  def limit(value, range):
      return scale(value, range, range)
  end


  rq_init_comm_if_connected(9, "1")
  rq_init_comm_if_connected(2, "2")
  rq_init_comm_if_connected(3, "3")
  rq_init_comm_if_connected(4, "4")
  rq_print_connected_grippers()
  rq_gripper_communication_thread = run rq_gripper_communication()
  set_closed_norm(97.6470588235294, 1)
  set_open_norm(1.1764705882352942, 1)
  set_closed_mm(0.0, 1)
  set_open_mm(53.0, 1)
  set_closed_norm(100.0, 2)
  set_open_norm(0.0, 2)
  set_closed_mm(0.0, 2)
  set_open_mm(50.0, 2)
  set_closed_norm(100.0, 3)
  set_open_norm(0.0, 3)
  set_closed_mm(0.0, 3)
  set_open_mm(50.0, 3)
  set_closed_norm(100.0, 4)
  set_open_norm(0.0, 4)
  set_closed_mm(0.0, 4)
  set_open_mm(50.0, 4)
  rq_current_limit_enabled = False
  while(not rq_gripper_communication_thread_started):
      sync()
  end
  # end: URCap Installation Node
  # begin: URCap Installation Node
  #   Source: OPC UA, 2.0.2, Rocketfarm AS
  #   Type: OPC UA
  global opcua_daemon = rpc_factory("xmlrpc", "http://127.0.0.1:40409/RPC2")
  def opcua_client_connect(address):
  return opcua_daemon.client_connect(address)
  end
  def opcua_client_get_id(client_name):
  return opcua_daemon.client_get_id(client_name)
  end
  def opcua_client_try_connect(client_id):
  opcua_result = False
  if (opcua_daemon.client_connect(client_id)):
  sleep(0.01)
  opcua_result = opcua_daemon.client_is_connected(client_id)
  opcua_retry = 10
  while ( (not opcua_result) and (opcua_retry > 0) ):
  sleep(0.1)
  opcua_result = opcua_daemon.client_is_connected(client_id)
  opcua_retry = opcua_retry - 1
  end
  end
  return opcua_result
  end
  def opcua_client_disconnect(client_id):
  return opcua_daemon.client_disconnect(client_id)
  end
  def opcua_client_is_connected(client_id):
  return opcua_daemon.client_is_connected(client_id)
  end
  def opcua_client_read_byid(client_id, namespace_id, variable_id):
  return opcua_daemon.client_read_variable_by_id(client_id, namespace_id, variable_id)
  end
  def opcua_client_read_byname(client_id, namespace_id, variable_name):
  return opcua_daemon.client_read_variable_by_name(client_id, namespace_id, variable_name)
  end
  def opcua_client_write_byid(client_id, namespace_id, variable_id, variable_value):
  return opcua_daemon.client_write_variable_by_id(client_id, namespace_id, variable_id, variable_value)
  end
  def opcua_client_write_byname(client_id, namespace_id, variable_name, variable_value):
  return opcua_daemon.client_write_variable_by_name(client_id, namespace_id, variable_name, variable_value)
  end
  def opcua_client_last_error(client_id):
  return opcua_daemon.client_get_last_error(client_id)
  end
  def opcua_server_read_byname(variable_name):
  return opcua_daemon.server_read_variable_by_name(variable_name)
  end
  def opcua_server_write_byname(variable_name, variable_value):
  return opcua_daemon.server_write_variable_by_name(variable_name, variable_value)
  end
  def opcua_server_last_error():
  return opcua_daemon.server_get_last_error()
  end
  def opcua_error_to_string(errorCode):
  return opcua_daemon.error_code_to_string(errorCode)
  end
  # end: URCap Installation Node
  step_count_7be696b6_0fa4_4b27_b09b_633ea860953e = 0.0
  thread Step_Counter_Thread_93e352b0_e34b_423c_bc3a_28ecb8afdc0a():
    while (True):
      step_count_7be696b6_0fa4_4b27_b09b_633ea860953e = step_count_7be696b6_0fa4_4b27_b09b_633ea860953e + 1.0
      sync()
    end
  end
  run Step_Counter_Thread_93e352b0_e34b_423c_bc3a_28ecb8afdc0a()
  global AMR_Position=struct(position_identifier=0, x1=0, x2=0, y1=0, y2=0, theta1=0, theta2=0)
  global CAM_Pose=p[0,0,0,0,0,0]
  global CAM_Relation=""
  global CMD_Abort=  False
  global CMD_Clear=  False
  global CMD_Reset=  False
  global CMD_Start=  False
  global CMD_Suspend=  False
  global CMD_Unhold=  False
  global CMD_Unsuspend=  False
  global CNT_Rack_Output=0
  global FNC_Freedrive=  False
  global PRC_TubCounter=0
  global PRC_TubNumber=0
  global STP=0
  global easyPickCount=0
  global easyPickCount_5=0
  global easyPickNoObj=0
  global easyPickNoObj_5=0
  global easyPickParts=0
  global easyPickParts_5=0
  global TMR_Barcode=0
  global Container_mid_1_p=p[-.379239199143, -.127191311915, .299999999998, .000000000046, -.000000000021, -1.247199999994]
  global Container_mid_1_q=[-2.477408934449926, -1.2969853503591224, -1.875639182904262, -1.539621866126728, 1.5731943360401213, -2.8009955944022717]
  global Container_capt_p=p[-.525590029047, .407247642794, .411588185841, -.000000000107, .000000000065, -2.896148821900]
  global Container_capt_q=[-3.5968351615224767, -2.0050156108707204, -0.8176271154495112, -1.8895759482008394, 1.5730967555598792, -2.2743681102957645]
  global Waypoint_6_p=p[.008800512419, -.547926542621, .402696567415, -.589884378425, -.007228654778, -.061268144704]
  global Waypoint_6_q=[-1.2044575850116175, -1.3416667741588135, -1.8272563219070435, -0.9884541195682068, 1.3621035814285278, -2.7712565104113978]
  global Waypoint_18_p=p[-.178371829612, -.433927395311, .368082383916, -.086593488055, .704679941724, -.007869906074]
  global Waypoint_18_q=[-1.265390698109762, -1.3355963987163086, -1.7944865226745605, -1.7402602634825648, 0.8780410885810852, -2.7713127771960657]
  global Waypoint_12_p=p[.008800512419, -.547926542621, .402696567415, -.589884378425, -.007228654778, -.061268144704]
  global Waypoint_12_q=[-1.2044575850116175, -1.3416667741588135, -1.8272563219070435, -0.9884541195682068, 1.3621035814285278, -2.7712565104113978]
  global Waypoint_19_p=p[-.178371829612, -.433927395311, .368082383916, -.086593488055, .704679941724, -.007869906074]
  global Waypoint_19_q=[-1.265390698109762, -1.3355963987163086, -1.7944865226745605, -1.7402602634825648, 0.8780410885810852, -2.7713127771960657]
  global Vial_above_p=p[.017105793010, -.652093028359, .184920586844, .000000000272, .000000000270, 1.564063451276]
  global Vial_above_q=[-1.3375440709712851, -1.9618096977868804, -1.4665759083780685, -1.2837941559171444, 1.5732503672317195, -4.47276330421513]
  global Vial_pick_point_p=p[.017105792852, -.648922724010, .093307568731, .000000000271, .000000000270, 1.564063451276]
  global Vial_pick_point_q=[-1.3366329456391917, -2.0375277831965413, -1.6071432798879028, -1.0675084332049813, 1.57309887265915, -4.471135348858068]
  global Waypoint_20_p=p[.019227646885, -.648669633640, .184920586950, .000000000000, .000000000000, .024063451426]
  global Waypoint_20_q=[-1.3331129109407733, -1.9540750545686123, -1.4775914902901128, -1.280581784992414, 1.5733500744865856, -2.928303704452631]
  global Waypoint_33_p=p[-.032361834699, -.348336136197, .391475576335, -.000008499254, .000014589902, -.004651426820]
  global Waypoint_33_q=[-1.2709335019096129, -1.1914598663441005, -1.708995335060501, -1.8117888533498316, 1.5729683532263925, -2.8379347397710237]
  global Vial_3FG_place_p=p[-.031858676359, -.349402499566, .145301120695, .000000000000, .000000000000, .000000000000]
  global Vial_3FG_place_q=[-1.2723975525801707, -1.252376585823825, -2.3128114007049496, -1.1470592278900167, 1.5730548099411423, -2.8414815174610535]
  global Waypoint_34_p=p[-.032361834699, -.348336136197, .391475576335, -.000008499254, .000014589902, -.004651426820]
  global Waypoint_34_q=[-1.2709335019096129, -1.1914598663441005, -1.708995335060501, -1.8117888533498316, 1.5729683532263925, -2.8379347397710237]
  global cap_dump_p=p[-.139168676487, -.420163541420, .146096395183, .000000000000, .000000000000, .000000000000]
  global cap_dump_q=[-1.584588644510994, -1.5093464179777323, -2.1118449369620347, -1.091059703602438, 1.5728943834877336, -3.154014906686923]
  global Waypoint_35_p=p[-.032361834699, -.348336136197, .391475576335, -.000008499254, .000014589902, -.004651426820]
  global Waypoint_35_q=[-1.2709335019096129, -1.1914598663441005, -1.708995335060501, -1.8117888533498316, 1.5729683532263925, -2.8379347397710237]
  global Waypoint_36_p=p[-.032361834699, -.348336136197, .391475576335, -.000008499254, .000014589902, -.004651426820]
  global Waypoint_36_q=[-1.2709335019096129, -1.1914598663441005, -1.708995335060501, -1.8117888533498316, 1.5729683532263925, -2.8379347397710237]
  global Waypoint_37_p=p[-.032361834699, -.348336136197, .391475576335, -.000008499254, .000014589902, -.004651426820]
  global Waypoint_37_q=[-1.2709335019096129, -1.1914598663441005, -1.708995335060501, -1.8117888533498316, 1.5729683532263925, -2.8379347397710237]
  global Vial_liq_above_p=p[-.025303660977, -.338758622354, .426628485936, -1.315858642253, .800043520260, -.928295855026]
  global Vial_liq_above_q=[-0.3789628187762659, -1.5149522957256814, -2.263045310974121, 0.7870649534412841, -0.750984017048971, -3.2237566153155726]
  global Vial_liq_pick_1_p=p[-.002660428945, -.335984893034, .159389832934, -1.150456778400, .673175527684, -1.010612657503]
  global Vial_liq_pick_1_q=[-0.3660772482501429, -1.4503649038127442, -2.4056053161621094, -1.994692941705221, 0.8039668202400208, -0.2508929411517542]
  global Vial_liq_pick_2_p=p[-.041402486291, -.356791603314, .125395323246, -1.143483969075, .651070210027, -.878721885453]
  global Vial_liq_pick_2_q=[-0.4426233705502476, -1.437252121513727, -2.551930962114307, -1.776528229806984, 0.6562026234073748, -0.43018811960029524]
  global Liquid_midway_p=p[.057575295009, -.583081747994, .306414980749, -1.351675548728, .120935756539, -.096908606303]
  global Liquid_midway_q=[-0.895174805318014, -1.7035466633238734, -2.380953073501587, 0.631549521083496, 0.7706599235534668, -2.9455552736865442]
  global shake_1_p=p[.057574880217, -.583085370269, .306422893466, -1.360996190983, -.155555042453, -.438136255921]
  global shake_1_q=[-0.8951800505267542, -1.7035466633238734, -2.380937099456787, 0.6315542894550782, 0.7706599235534669, -2.5394540616517496]
  global shake_2_p=p[.057581636113, -.583090570002, .306439684073, -1.308767904323, .368530312677, .214926493520]
  global shake_2_q=[-0.8951714674579065, -1.7035395107665003, -2.380906343460083, 0.6315504747578125, 0.7706480026245118, -3.3161255787892268]
  global drop_above_1_p=p[.268235025993, -.467784390499, .226219872376, -1.027832627524, -.430841408251, 1.004603115937]
  global drop_above_1_q=[-0.935645882283346, -1.6663371525206507, -2.4252893924713135, 0.41966931402172847, 1.8470635414123535, -3.4600217978106897]
  global drop_above_2_p=p[.219042229014, -.470775657081, .133754190740, -.313004595901, -.344395319364, 1.500564994056]
  global drop_above_2_q=[-1.0601594887284795, -1.70046459045642, -2.0799996233759863, -0.7243227230676759, 1.9429634314685202, -4.115129153870795]
  global liq_tran_1_p=p[.213067510942, -.469567035397, .100231043184, .251862243732, .217902579404, 1.592812335393]
  global liq_tran_1_q=[-0.7789645168037476, -1.822364827406652, -1.8643518410805573, -1.252158963840138, 1.3768134449520435, -3.9328333233290254]
  global Waypoint_21_p=p[.187119460405, -.493959476151, .133754190608, -.313004596540, -.344395317757, 1.500564993991]
  global Waypoint_21_q=[-1.1418328121400876, -1.7310553375189475, -2.033634768766424, -0.772026910513711, 1.958578934631971, -4.201588449364511]
  global liq_tran_2_p=p[.195957706507, -.493022614126, .100231042689, .160718757180, .109807038912, 1.525321508623]
  global liq_tran_2_q=[-0.881740380645474, -1.8244526267589851, -1.865100964490387, -1.1608866323693583, 1.4631433601076713, -3.973915130363038]
  global Vial_drop_above_p=p[.000324902251, -.648569523142, .221894115667, -.873462921366, 1.165852672573, -1.482720593185]
  global Vial_drop_above_q=[-1.0576906334721352, -2.393016994184633, -0.9236232851859159, -2.5729213042279273, 0.7903331288549689, -0.33286325848155585]
  global Vial_liq_drop_p=p[.001020867953, -.647659915585, .092915870838, -.834762611599, 1.081942994823, -1.540647900176]
  global Vial_liq_drop_q=[-1.0631954168193474, -2.4447642951220825, -1.128811017825127, -2.1983115491972294, 0.8130148661460634, -0.38984988696911316]
  global Waypoint_9_p=p[.206300564882, -.401796282405, .209941275233, .000000000049, .000000000063, 1.560839127857]
  global Waypoint_9_q=[-0.7963359454512808, -1.4686025034365713, -1.9726632321075135, -1.2709582822971974, 1.5730203818053559, -3.9272300959189193]
  global Waypoint_10_p=p[.200865824304, -.400817692024, .105072686738, .000000000049, .000000000061, 1.560839127855]
  global Waypoint_10_q=[-0.8042914374275529, -1.5824702465090397, -2.1630314773482997, -0.9667217216455377, 1.5726337265768082, -3.9342465798801403]
  global Waypoint_11_p=p[.200865824280, -.400817691999, .325177251663, .000000000049, .000000000061, 1.560839127855]
  global Waypoint_11_q=[-0.8031609769098491, -1.4190566846320642, -1.7173307870816634, -1.5758364190022327, 1.5730457436482617, -3.935202548332848]
  global Waypoint_7_p=p[-.615828862681, .233809157513, .299999999960, .005115849907, .008741794022, -2.111813105778]
  global Waypoint_7_q=[-3.2957401409809868, -1.9361965884744503, -1.2056078493731617, -1.569266158150004, 1.5650998100608482, -2.7562028470627613]
  global Waypoint_8_p=p[-.615828862366, .233809157463, .013910424379, .005115849905, .008741794020, -2.111813105780]
  global Waypoint_8_q=[-3.2964782505943173, -2.1586184138220776, -1.6500090431308791, -0.9024541777239836, 1.5648120752692236, -2.7547026290098384]
  global Waypoint_13_p=p[-.479450777041, .284140798427, .125270103493, -.276792173670, 2.098433187455, -2.121256516887]
  global Waypoint_13_q=[-2.8915050665484827, -1.9549266300597132, -2.2318272590637207, -1.6654960117735804, 0.020810842514038086, -0.4019392172442835]
  global Waypoint_70_p=p[-.472820924464, .292439826304, .207418370234, -.259787347864, -2.053484648504, 2.070709755662]
  global Waypoint_70_q=[-2.969927421603815, -2.07168115810532, -1.6835546062719366, -2.4953958198513964, 0.4489790927922641, -0.005578998612037367]
  global Waypoint_1_p=p[-.312961047461, -.152991312519, .223609826854, -.745314530454, -1.713873240489, 1.673341715282]
  global Waypoint_1_q=[-2.3560472170459192, -2.183784624139303, -1.4583134651184082, -2.6435262165465296, 1.6522362232208252, 0.043451953679323196]
  global Waypoint_16_p=p[-.113749865836, -.390110151572, .317307487562, -.519383711706, -.839884211339, 1.756868173041]
  global Waypoint_16_q=[-1.8909733931170862, -1.720626016656393, -1.5115610361099243, -2.1240560017027796, 2.1809096336364746, 0.7227501273155212]
  global Waypoint_15_p=p[.029144035010, -.436802470887, .327885032028, -.521560953301, -.623641814548, 1.862659450154]
  global Waypoint_15_q=[-1.564817253743307, -1.556895188321807, -1.6826975345611572, -1.6944714985289515, 2.2362685203552246, 1.117417335510254]
  global Waypoint_14_p=p[.068712235638, -.569419545175, .285215357659, -.679242949116, -.712065334485, 1.394044574094]
  global Waypoint_14_q=[-1.5731792953485346, -1.8029235103747094, -1.6781008808776736, -1.2218450646111982, 2.4719572998240125, 1.6394218026856375]
  global Waypoint_17_p=p[-.047220457210, -.557624911767, .136370962514, -.679242949107, -.712065334475, 1.394044574096]
  global Waypoint_17_q=[-1.7740079055958748, -2.0023561428872334, -1.7577251142892676, -1.18903287716154, 2.4487287370345143, 1.322902469273079]
  global Waypoint_25_p=p[.065436479647, -.569388431626, .287820755049, -.679242949185, -.712065334557, 1.394044574070]
  global Waypoint_25_q=[-1.5789263550890595, -1.8020194754825436, -1.6702557537748035, -1.237882536889547, 2.471995808083492, 1.6301087487321393]
  global Waypoint_73_p=p[.200650292861, -.570238752026, .330084459991, 1.360500825815, .021700154388, 2.681649888469]
  global Waypoint_73_q=[-0.7671117850166942, -2.170180210127774, -0.8654875324671831, -2.4760661058854714, 1.019668964673781, 1.1886838746103445]
  global Waypoint_51_p=p[.143029822311, -.569853361759, .275754213782, 1.297896664289, .026410127072, 2.712872144875]
  global Waypoint_51_q=[-0.8339941389801577, -2.0499669090260237, -1.181859109742545, -2.1992567984298894, 0.9933974691724003, 1.1053015960835664]
  global Waypoint_55_p=p[.073857253409, -.577012553496, .221504790513, 1.297896665457, .026410123899, 2.712872144362]
  global Waypoint_55_q=[-0.9235026509638331, -2.0031911550113533, -1.4013130080059835, -1.9791459123699324, 0.9364696407276547, 1.0224867664664226]
  global Waypoint_56_p=p[.135677267144, -.579447716527, .242231366835, 1.555421348248, .015405426287, 2.555899922373]
  global Waypoint_56_q=[-0.8277598345563266, -2.1783820448240228, -1.1390951780517948, -2.3437042464770936, 0.9222576608739947, 1.2572681804986878]
  global Waypoint_57_p=p[.143391004007, -.581808738942, .226065325532, 1.639743959545, .007914821713, 2.502360786858]
  global Waypoint_57_q=[-0.8163397121067408, -2.2409861865625498, -1.1056400409378426, -2.4000192569642436, 0.9131014133193622, 1.3141118037187605]
  global Waypoint_59_p=p[.272401132286, -.578182925380, .239561357365, 2.126997331910, .113921148153, 2.155615020515]
  global Waypoint_59_q=[-0.6600120703326624, -2.700596948663229, -0.4450863301753998, -3.1158048115172328, 0.9327830672264099, 1.686402678489685]
  global Waypoint_58_p=p[.223648508176, -.578477552733, .276546452136, 2.174288010107, -.044108754041, 2.058653287678]
  global Waypoint_58_q=[-0.7290484882560344, -2.6749849159411134, -0.44426632073579775, -3.220833992584847, 0.9665895014735898, 1.686536774549042]
  global Waypoint_60_p=p[-.013316432876, -.544772031582, .383371643081, 2.208233379808, .037543335712, 2.097559881761]
  global Waypoint_60_q=[-0.9328326161883087, -2.0999933666355775, -1.1958015693111372, -3.060905141293654, 0.690378518537611, 1.7121940951337198]
  global Waypoint_61_p=p[-.412188693372, -.356446875193, .383371643081, 1.751740964455, -.739956256289, 1.600691174920]
  global Waypoint_61_q=[-1.766185342973321, -2.0999933666355775, -1.1958015693111372, -3.060905141293654, 0.690378518537611, 1.7121940951337198]
  global Waypoint_62_p=p[-.542658707241, -.114281911009, .251261544113, 1.813043609523, -.679411528034, 1.655271622964]
  global Waypoint_62_q=[-2.158300033470912, -1.9418836862428677, -1.8142999147147894, -2.778920736683023, 0.21900622104017292, 1.8983390235012934]
  global Waypoint_63_p=p[-.532496162227, -.127810170801, .159342327524, 1.813043609478, -.679411528027, 1.655271622994]
  global Waypoint_63_q=[-2.1232624524640213, -2.086114053133292, -1.8911847933380095, -2.5248779786918614, 0.2536249317365024, 1.864405460969639]
  global Waypoint_52_p=p[-.576034890047, -.066269986912, .306739617770, .862065193359, -.255405331227, 2.195240951653]
  global Waypoint_52_q=[-2.4808268779922003, -1.5303848711262056, -1.876845562237385, -1.1257011427858359, 0.8740163290385958, -0.15002503295170655]
  global Waypoint_69_p=p[-.581965326699, -.059291422286, .312082125679, .862065195757, -.255405329473, 2.195240950921]
  global Waypoint_69_q=[-2.500621389999687, -1.5361955180345959, -1.8614018767844556, -1.1190332887072278, 0.8777181708365909, -0.17540933674578696]
  global Waypoint_71_p=p[-.581965326670, -.059291422265, .290575803625, .862065195756, -.255405329472, 2.195240950921]
  global Waypoint_71_q=[-2.5007210652259566, -1.5510704265538795, -1.9040561970342402, -1.0615823481403304, 0.8776641555740685, -0.17528706367848557]
  global Waypoint_72_p=p[-.581965326627, -.059291422244, .350142125738, 1.757497900770, -.677813691618, 1.696469016977]
  global Waypoint_72_q=[-2.3014470577960933, -1.774776476208789, -1.7081605706825291, -2.8433626113276596, 0.07508598567825443, 1.682946898281932]
  global Waypoint_68_p=p[-.333292906431, -.480744165508, .350142125738, 2.217519979286, .140864133573, 2.209123277630]
  global Waypoint_68_q=[-1.438387057796029, -1.774776476208789, -1.7081605706825291, -2.8433626113276596, 0.07508598567825443, 1.682946898281932]
  global TMR_Barcode_is_counting=False
  thread Timer_Thread():
    while (True):
      if (TMR_Barcode_is_counting):
        TMR_Barcode = TMR_Barcode + get_steptime()
      end
      sync()
    end
  end
  run Timer_Thread()
  def Sub_Vision_V18():
    $ 697 "Sub_Vision_V18" "noBreak"
    $ 698 "PreSettings"
    $ 699 "CAM_LM_Detected≔ False "
    global CAM_LM_Detected=  False
    $ 700 "CAM_Captures≔0"
    global CAM_Captures=0
    $ 701 "CAM_Pose≔p[0,0,0,0,0,0]"
    global CAM_Pose=p[0,0,0,0,0,0]
    $ 702 "CAM_LM_Refinmnt≔ False "
    global CAM_LM_Refinmnt=  False
    $ 703 "CAM_LM_Refined≔ False "
    global CAM_LM_Refined=  False
    $ 704 "CAM_LM_Deviatn≔p[0,0,0,0,0,0]"
    global CAM_LM_Deviatn=p[0,0,0,0,0,0]
    $ 705 "CAM_LM_ID≔0"
    global CAM_LM_ID=0
    $ 706 "CAM_Done≔ False "
    global CAM_Done=  False
    $ 707 "CAM_CNT_Obj≔0"
    global CAM_CNT_Obj=0
    $ 708 "CAM_Result = []"
    CAM_Result = []
    $ 709 "OBJ_Detected≔ False "
    global OBJ_Detected=  False
    $ 710 "FRM_Reference≔p[0,0,0,0,0,0]"
    global FRM_Reference=p[0,0,0,0,0,0]
    $ 711 "'=========='"
    # '=========='
    $ 712 "Switch Action"
    switch_1 = Action
    $ 713 "Case 13"
    if (13 == switch_1):
    elif (15 == switch_1):
      $ 831 "Case 15"
    elif (131 == switch_1):
      $ 877 "Case 131"
      $ 878 "Read (SensoPart)"
      $ 879 "Action_Info≔'search for landmark'"
      global Action_Info="search for landmark"
      $ 880 "CAM_LM≔CAM_LMs[4]"
      global CAM_LM=CAM_LMs[4]
      $ 881 "CAM_Relation≔CAM_LM.capture_relation"
      global CAM_Relation=CAM_LM.capture_relation
      $ 882 "go to capture pose"
      $ 885 "If ITM_ID≟1 and JIG≟7"
      if (ITM_ID == 1  and  JIG == 7):
        $ 886 "PSE_T≔uLM_Cap_SSRack"
        global PSE_T=uLM_Cap_SSRack
      else:
        $ 887 "ElseIf ITM_ID≟5 and JIG≟7"
        if (ITM_ID == 5  and  JIG == 7):
          $ 888 "PSE_T≔FRM_Cap_SSRack"
          global PSE_T=FRM_Cap_SSRack
        else:
          $ 889 "ElseIf ITM_ID≟13 and JIG≟7"
          if (ITM_ID == 13  and  JIG == 7):
            $ 890 "PSE_T≔FRM_pick_rack_const"
            global PSE_T=p[-0.5568395192387274,0.34423986364170267,0.44698620470146266,-1.0069110132199915E-6,3.378712467497258E-5,-8.002029546773325E-6]
          else:
            $ 891 "ElseIf ITM_ID≟1 and JIG≟15"
            if (ITM_ID == 1 and JIG == 15):
              $ 892 "MoveJ"
              $ 893 "Container_mid_1" "breakAfter"
              movej(get_inverse_kin(Container_mid_1_p, qnear=Container_mid_1_q), a=1.3962634015954636, v=1.0471975511965976, r=0.05)
              $ 894 "Container_capt" "breakAfter"
              movej(get_inverse_kin(Container_capt_p, qnear=Container_capt_q), a=1.3962634015954636, v=1.0471975511965976)
              $ 895 "PSE_T≔FRM_Container_S_const"
              global PSE_T=p[-0.510412665574981,0.40064363362973565,0.41159789496794374,-1.1370875604168537E-5,-3.643547521609506E-6,-2.896122366208473]
            end
          end
        end
      end
      $ 896 "do_transition(PSE_T, keep_rxry=False)"
      do_transition(PSE_T, keep_rxry=False)
      $ 897 "Set"
      set_tcp(p[0.0,0.0,0.161,3.1415,0.0,0.0])
      $ 898 "MoveJ"
      $ 899 "PSE_T" "breakAfter"
      movej(PSE_T, a=1.3962634015954636, v=1.7453292519943295)
      $ 900 "CAM_Pose≔get_actual_tcp_pose()"
      global CAM_Pose= get_actual_tcp_pose ()
      $ 901 "Loop  not CAM_Done and  not ERROR.FLAG and  not CMD_Stop"
      while (  not  CAM_Done  and    not  ERROR.FLAG  and    not  CMD_Stop):
        $ 902 "adjust capture pose"
        $ 903 "If CAM_LM_Detected and CAM_LM_Refinmnt"
        if (CAM_LM_Detected  and  CAM_LM_Refinmnt):
          $ 904 "PSE_T≔p[0,0,0.300,0,0,0]"
          global PSE_T=p[0,0,0.300,0,0,0]
          $ 905 "CAM_Pose≔PSE_T"
          global CAM_Pose=PSE_T
          $ 906 "If  not is_reachable(FRM_Reference,[PSE_T])"
          if (  not  is_reachable(FRM_Reference,[PSE_T])):
            $ 907 "Error"
            $ 908 "set_error(ERROR_POSE_NOT_REACHABLE)"
            set_error(ERROR_POSE_NOT_REACHABLE)
          end
          $ 909 "If  not ERROR.FLAG"
          if (  not  ERROR.FLAG):
            $ 910 "MoveJ"
            $ 911 "PSE_T" "breakAfter"
            set_tcp(p[0.0,0.0,0.161,0.0,0.0,0.0])
            movej(pose_trans(FRM_Reference, PSE_T), a=0.8726646259971648, v=1.3962634015954636)
            $ 912 "CAM_LM_Refined≔ True "
            global CAM_LM_Refined=  True
          end
        else:
          $ 913 "ElseIf  not CAM_LM_Detected and CAM_Captures>0"
          if (  not  CAM_LM_Detected  and  CAM_Captures>0):
            $ 914 "MoveL"
            $ 915 "If FRM_Reference≟p[0,0,0,0,0,0]"
            if (FRM_Reference == p[0,0,0,0,0,0]):
              $ 916 "PSE_T≔get_random_pose(pose_ref=CAM_Pose, mode='cubic', range_max=[0.150,0.150,0.015])"
              global PSE_T=get_random_pose(pose_ref=CAM_Pose, mode="cubic", range_max=[0.150,0.150,0.015])
            else:
              $ 921 "Else" "noBreak"
              $ 922 "PSE_T≔get_random_pose(pose_ref=CAM_Pose, mode='rotation', range_max=[10,10,0])"
              global PSE_T=get_random_pose(pose_ref=CAM_Pose, mode="rotation", range_max=[10,10,0])
              $ 923 "CAM_LM_Refined≔ True "
              global CAM_LM_Refined=  True
            end
            $ 924 "If get_inverse_kin_has_solution(pose_trans(FRM_Reference, PSE_T))"
            if (get_inverse_kin_has_solution( pose_trans (FRM_Reference, PSE_T))):
              $ 925 "Comment"
              # Comment
              $ 926 "PSE_T" "breakAfter"
              set_tcp(p[0.0,0.0,0.161,3.1415,0.0,0.0])
              movel(pose_trans(FRM_Reference, PSE_T), a=0.03, v=0.05)
            else:
              $ 927 "Else" "noBreak"
              $ 928 "'If random pose is out of reach, set the initial cam pose'"
              # 'If random pose is out of reach, set the initial cam pose'
              $ 929 "PSE_T≔CAM_Pose"
              global PSE_T=CAM_Pose
            end
          end
        end
        $ 930 "Wait: 2.0"
        sleep(2.0)
        $ 931 "trigger"
        $ 932 "If ITM_ID≟1 and JIG≟7"
        if (ITM_ID == 1  and  JIG == 7):
          # begin: URCap Program Node
          #   Source: SensoPart VISOR Robotic, 2.0.0, SensoPart Industriesensorik GmbH
          #   Type: VISOR Trigger
          $ 933 "# 1 VISOR Trigger"
          visor_changeJob(1, "Landmark_INVITE_2", 6000)
          visor_trigger(1, 6000, "arm")
          # end: URCap Program Node
        else:
          $ 934 "ElseIf ITM_ID≟5 and JIG≟7"
          if (ITM_ID == 5  and  JIG == 7):
            # begin: URCap Program Node
            #   Source: SensoPart VISOR Robotic, 2.0.0, SensoPart Industriesensorik GmbH
            #   Type: VISOR Trigger
            $ 935 "# 1 VISOR Trigger"
            visor_changeJob(1, "Landmark_INVITE_2", 6000)
            visor_trigger(1, 6000, "arm")
            # end: URCap Program Node
          else:
            $ 936 "ElseIf ITM_ID≟13 and JIG≟7"
            if (ITM_ID == 13  and  JIG == 7):
              # begin: URCap Program Node
              #   Source: SensoPart VISOR Robotic, 2.0.0, SensoPart Industriesensorik GmbH
              #   Type: VISOR Trigger
              $ 937 "# 1 VISOR Trigger"
              visor_changeJob(1, "Landmark_INVITE_2", 6000)
              visor_trigger(1, 6000, "arm")
              # end: URCap Program Node
            else:
              $ 938 "ElseIf ITM_ID≟1 and JIG≟15"
              if (ITM_ID == 1 and JIG == 15):
                # begin: URCap Program Node
                #   Source: SensoPart VISOR Robotic, 2.0.0, SensoPart Industriesensorik GmbH
                #   Type: VISOR Trigger
                $ 939 "# 1 VISOR Trigger"
                visor_changeJob(1, "Container_S", 6000)
                visor_trigger(1, 6000, "arm")
                # end: URCap Program Node
              end
            end
          end
        end
        $ 943 "TM_3D_Found≔visor_partsFound(1)"
        global TM_3D_Found= visor_partsFound (1)
        $ 944 "If TM_3D_Found>0"
        if (TM_3D_Found>0):
          $ 945 "CAM_LM_Detected≔ True "
          global CAM_LM_Detected=  True
          $ 946 "CAM_Captures≔0"
          global CAM_Captures=0
        else:
          $ 947 "Else" "noBreak"
          $ 948 "CAM_LM_Detected≔ False "
          global CAM_LM_Detected=  False
          $ 949 "CAM_Captures≔CAM_Captures+1"
          global CAM_Captures=CAM_Captures+1
        end
        $ 954 "result"
        $ 955 "If CAM_LM_Detected"
        if (CAM_LM_Detected):
          $ 956 "If (CAM_LM_Refinmnt and CAM_LM_Refined) or  not CAM_LM_Refinmnt"
          if ((CAM_LM_Refinmnt  and  CAM_LM_Refined)  or    not  CAM_LM_Refinmnt):
            $ 1014 "If ITM_ID≟1 and JIG≟7"
            if (ITM_ID == 1  and  JIG == 7):
              $ 1015 "CAM_LM_SSRack≔visor_getPose3d(1, 0)"
              global CAM_LM_SSRack= visor_getPose3d (1, 0)
            else:
              $ 1016 "ElseIf ITM_ID≟5 and JIG≟7"
              if (ITM_ID == 5  and  JIG == 7):
                $ 1017 "CAM_LM_SSRack≔visor_getPose3d(1, 0)"
                global CAM_LM_SSRack= visor_getPose3d (1, 0)
              else:
                $ 1018 "ElseIf ITM_ID≟13 and JIG≟7"
                if (ITM_ID == 13  and  JIG == 7):
                  $ 1019 "CAM_LM_Bott≔visor_getPose3d(1, 0)"
                  global CAM_LM_Bott= visor_getPose3d (1, 0)
                else:
                  $ 1020 "ElseIf ITM_ID≟1 and JIG≟15"
                  if (ITM_ID == 1 and JIG == 15):
                    $ 1021 "CAM_LM_Cont_S≔visor_getPose3d(1, 0)"
                    global CAM_LM_Cont_S= visor_getPose3d (1, 0)
                  end
                end
              end
            end
            $ 1022 "CAM_Done≔ True "
            global CAM_Done=  True
          end
        else:
          $ 1023 "ElseIf  not CAM_LM_Detected and CAM_Captures<CAM_PRM_Retries"
          if (  not  CAM_LM_Detected  and  CAM_Captures<CAM_PRM_Retries):
            $ 1024 "CAM_LM_Refined≔ False "
            global CAM_LM_Refined=  False
          else:
            $ 1025 "ElseIf CAM_Captures≥CAM_PRM_Retries"
            if (CAM_Captures >= CAM_PRM_Retries):
              $ 1026 "CAM_Done≔ True "
              global CAM_Done=  True
              $ 1027 "Error"
              $ 1028 "set_error(ERROR_NO_LANDMARK)"
              set_error(ERROR_NO_LANDMARK)
            end
          end
        end
      end
    elif (151 == switch_1):
      $ 1029 "Case 151"
      $ 1030 "Detect (SensoPart)"
      $ 1031 "go to capture pose"
      $ 1032 "FRM_Reference≔FRM_Cap_SSRack"
      global FRM_Reference=FRM_Cap_SSRack
      $ 1033 "PSE_T≔p[0,0,-0.00,0,0,0]"
      global PSE_T=p[0,0,-0.00,0,0,0]
      $ 1034 "do_transition(pose_trans(FRM_Reference, PSE_T), keep_rxry=False)"
      do_transition( pose_trans (FRM_Reference, PSE_T), keep_rxry=False)
      $ 1035 "JNT_Q≔get_actual_joint_positions()"
      global JNT_Q= get_actual_joint_positions ()
      $ 1036 "JNT_Q≔[JNT_Q[0], JNT_Q[1], JNT_Q[2], JNT_Q[3], JNT_Q[4], 0]"
      global JNT_Q=[JNT_Q[0], JNT_Q[1], JNT_Q[2], JNT_Q[3], JNT_Q[4], 0]
      $ 1037 "Set"
      set_tcp(p[0.0,0.0,0.161,3.1415,0.0,0.0])
      $ 1038 "movej(get_inverse_kin(pose_trans(FRM_Reference, PSE_T), qnear=JNT_Q))"
      movej(get_inverse_kin( pose_trans (FRM_Reference, PSE_T), qnear=JNT_Q))
      $ 1039 "CAM_Pose≔pose_trans(pose_inv(FRM_Reference), get_actual_tcp_pose())"
      global CAM_Pose= pose_trans ( pose_inv (FRM_Reference),  get_actual_tcp_pose ())
      $ 1040 "Loop  not CAM_Done and  not ERROR.FLAG and  not CMD_Stop"
      while (  not  CAM_Done  and    not  ERROR.FLAG  and    not  CMD_Stop):
        $ 1041 "If  not OBJ_Detected and CAM_Captures>0"
        if (  not  OBJ_Detected  and  CAM_Captures>0):
          $ 1042 "MoveL"
          $ 1043 "If FRM_Reference≟p[0,0,0,0,0,0]"
          if (FRM_Reference == p[0,0,0,0,0,0]):
            $ 1045 "PSE_T≔get_random_pose(pose_ref=CAM_Pose, mode='rotation', range_max=[15,15,0])"
            global PSE_T=get_random_pose(pose_ref=CAM_Pose, mode="rotation", range_max=[15,15,0])
          else:
            $ 1046 "Else" "noBreak"
            $ 1047 "PSE_T≔get_random_pose(pose_ref=CAM_Pose, mode='rotation', range_max=[10,10,0])"
            global PSE_T=get_random_pose(pose_ref=CAM_Pose, mode="rotation", range_max=[10,10,0])
          end
          $ 1048 "If get_inverse_kin_has_solution(pose_trans(FRM_Reference, PSE_T))"
          if (get_inverse_kin_has_solution( pose_trans (FRM_Reference, PSE_T))):
            $ 1049 "PSE_T" "breakAfter"
            set_tcp(p[0.0,0.0,0.161,3.1415,0.0,0.0])
            movel(pose_trans(FRM_Reference, PSE_T), a=0.03, v=0.05)
          else:
            $ 1050 "Else" "noBreak"
            $ 1051 "'If random pose is out of reach, set the initial cam pose'"
            # 'If random pose is out of reach, set the initial cam pose'
            $ 1052 "PSE_T≔CAM_Pose"
            global PSE_T=CAM_Pose
            $ 1053 "PSE_T" "breakAfter"
            set_tcp(p[0.0,0.0,0.161,3.1415,0.0,0.0])
            movel(pose_trans(FRM_Reference, PSE_T), a=0.03, v=0.05)
          end
        end
        $ 1054 "Wait: 0.5"
        sleep(0.5)
        $ 1055 "Set"
        set_tcp(p[0.0,0.0,0.161,3.1415,0.0,0.0])
        # begin: URCap Program Node
        #   Source: SensoPart VISOR Robotic, 2.0.0, SensoPart Industriesensorik GmbH
        #   Type: VISOR Trigger
        $ 1056 "# 1 VISOR Trigger"
        visor_changeJob(1, "Object Detection Single", 6000)
        visor_trigger(1, 6000, "arm")
        # end: URCap Program Node
        $ 1057 "If visor_isResponseOk(1)"
        if ( visor_isResponseOk (1)):
          $ 1058 "CAM_CNT_Obj≔visor_partsFound(1)"
          global CAM_CNT_Obj= visor_partsFound (1)
          $ 1059 "CAM_OBJ_Pose≔visor_getPose3d(1, 0)"
          global CAM_OBJ_Pose= visor_getPose3d (1, 0)
          $ 1060 "If CAM_CNT_Obj>0"
          if (CAM_CNT_Obj>0):
            $ 1061 "CAM_OBJ_Color≔visor_getAdditionalData(1, 0)"
            global CAM_OBJ_Color= visor_getAdditionalData (1, 0)
            $ 1062 "CAM_DetectScore≔to_num(visor_getAdditionalData(1, 1))/1000"
            global CAM_DetectScore=to_num( visor_getAdditionalData (1, 1))/1000
            $ 1063 "OBJ_Detected≔ True "
            global OBJ_Detected=  True
          end
        else:
          $ 1064 "Else" "noBreak"
          $ 1065 "CAM_Captures≔CAM_Captures+1"
          global CAM_Captures=CAM_Captures+1
        end
        $ 1066 "If OBJ_Detected"
        if (OBJ_Detected):
          $ 1067 "Get object data"
          $ 1068 "PRC_CntDetect≔0"
          global PRC_CntDetect=0
          $ 1069 "Loop PRC_CntDetect<CAM_CNT_Obj"
          while (PRC_CntDetect<CAM_CNT_Obj):
            $ 1070 "get object and jig number"
            $ 1071 "If ITM_ID≟1 and JIG≟7"
            if (ITM_ID == 1  and  JIG == 7):
              $ 1072 "FRM_Reference≔FRM_Cap_SSRack"
              global FRM_Reference=FRM_Cap_SSRack
            else:
              $ 1073 "ElseIf ITM_ID≟5 and JIG≟7"
              if (ITM_ID == 5  and  JIG == 7):
                $ 1074 "FRM_Reference≔uLM_Cap_SSRack"
                global FRM_Reference=uLM_Cap_SSRack
              end
            end
            $ 1077 "PSE_T≔pose_trans(pose_inv(FRM_Reference), CAM_OBJ_Pose)"
            global PSE_T= pose_trans ( pose_inv (FRM_Reference), CAM_OBJ_Pose)
            $ 1078 "CAM_Result.append(get_pattern_counter(PSE_T, 'X', pattern=[10, 5], patternsize=[0.181, 0.081]))"
            CAM_Result.append(get_pattern_counter(PSE_T, "X", pattern=[10, 5], patternsize=[0.181, 0.081]))
            $ 1079 "PRC_CntDetect≔PRC_CntDetect+1"
            global PRC_CntDetect=PRC_CntDetect+1
          end
          $ 1080 "CAM_Done≔ True "
          global CAM_Done=  True
        else:
          $ 1081 "ElseIf CAM_Captures≥CAM_PRM_Retries"
          if (CAM_Captures >= CAM_PRM_Retries):
            $ 1082 "CAM_Done≔ True "
            global CAM_Done=  True
          else:
            $ 1083 "Else" "noBreak"
            $ 1084 "CAM_Captures≔CAM_Captures+1"
            global CAM_Captures=CAM_Captures+1
          end
        end
      end
    end
    $ 1085 "'=========='"
    # '=========='
    $ 1086 "PostSettings"
    $ 1087 "FRM_Reference≔p[0,0,0,0,0,0]"
    global FRM_Reference=p[0,0,0,0,0,0]
    $ 1088 "Set"
    set_tcp(p[0.0,0.0,0.161,3.1415,0.0,0.0])
    $ 1089 "CAM_Pose≔p[0,0,0,0,0,0]"
    global CAM_Pose=p[0,0,0,0,0,0]
    $ 1090 "Action≔0"
    global Action=0
    $ 1091 "Action_Info≔''"
    global Action_Info=""
  end
  def Sub_AMR_MiR_V3():
    $ 1092 "Sub_AMR_MiR_V3" "noBreak"
    $ 1093 "PreSettings"
    $ 1094 "AMR_TargetList≔[1,2,3,4,5,21,22,23,24,31,32,33,34,35,36,37,38,41]"
    global AMR_TargetList=[1,2,3,4,5,21,22,23,24,31,32,33,34,35,36,37,38,41]
    $ 1095 "AMR_Done≔ False "
    global AMR_Done=  False
    $ 1096 "AMR_PosActual≔T2O_Current_Pos"
    global AMR_PosActual=modbus_get_signal_status("T2O_Current_Pos")
    $ 1097 "AMR_Attemps≔T2O_Nav_Attemps"
    global AMR_Attemps=modbus_get_signal_status("T2O_Nav_Attemps")
    $ 1098 "AMR_Battery≔MiR_Battery_Lvl"
    global AMR_Battery=modbus_get_signal_status("MiR_Battery_Lvl")
    $ 1099 "AMR_Charging≔(T2O_Charging≟1)"
    global AMR_Charging=(modbus_get_signal_status("T2O_Charging") == 1)
    $ 1100 "AMR_Position≔struct(position_identifier=T2O_Current_Pos, x1=MiR_Position_X1, x2=MiR_Position_X2, y1=MiR_Position_Y1, y2=MiR_Position_Y2, theta1=MiR_Theta_1, theta2=MiR_Theta_2) "
    global AMR_Position=struct(position_identifier=modbus_get_signal_status("T2O_Current_Pos"), x1=modbus_get_signal_status("MiR_Position_X1"), x2=modbus_get_signal_status("MiR_Position_X2"), y1=modbus_get_signal_status("MiR_Position_Y1"), y2=modbus_get_signal_status("MiR_Position_Y2"), theta1=modbus_get_signal_status("MiR_Theta_1"), theta2=modbus_get_signal_status("MiR_Theta_2"))
    $ 1101 "If MiR_Mode≠7"
    if (modbus_get_signal_status("MiR_Mode") != 7):
      $ 1102 "Error"
      $ 1103 "set_error(ERROR_AMR_WRONG_MODE)"
      set_error(ERROR_AMR_WRONG_MODE)
      $ 1104 "AMR_Done≔ True "
      global AMR_Done=  True
    end
    $ 1105 "'=========='"
    # '=========='
    $ 1106 "Switch STATE"
    switch_1 = STATE
    $ 1107 "Case 1"
    if (1 == switch_1):
      $ 1108 "stopping"
      $ 1109 "If T2O_Done≟1 and O2T_Acknowledge≟0"
      if (modbus_get_signal_status("T2O_Done") == 1  and  modbus_get_signal_status("O2T_Acknowledge") == 0):
        $ 1110 "Set O2T_Acknowledge=1"
        modbus_set_output_register("O2T_Acknowledge", 1)
      end
      $ 1111 "Set MiR_CMD_Stop=On"
      modbus_set_output_signal("MiR_CMD_Stop", True)
      $ 1112 "AMR_Position.position_identifier = 0"
      AMR_Position.position_identifier = 0
      $ 1113 "AMR_Done≔ True "
      global AMR_Done=  True
    elif (2 == switch_1):
      $ 1114 "Case 2"
      $ 1115 "stopped"
      $ 1116 "If MiR_State≠3 and MiR_State≠5"
      if (modbus_get_signal_status("MiR_State") != 3  and  modbus_get_signal_status("MiR_State") != 5):
        $ 1117 "Set MiR_CMD_Stop=Off"
        modbus_set_output_signal("MiR_CMD_Stop", False)
      end
    elif (3 == switch_1):
      $ 1118 "Case 3"
      $ 1119 "resetting"
      $ 1120 "Set O2T_Mis_Main=Off"
      modbus_set_output_signal("O2T_Mis_Main", False)
      $ 1121 "Set O2T_Mis_Charge=Off"
      modbus_set_output_signal("O2T_Mis_Charge", False)
      $ 1122 "If MiR_Mis_Queue>0"
      if (modbus_get_signal_status("MiR_Mis_Queue")>0):
        $ 1123 "Set MiR_CMD_Clear_Q=On"
        modbus_set_output_signal("MiR_CMD_Clear_Q", True)
        $ 1124 "Wait MiR_Mis_Queue≟0"
        while (not(modbus_get_signal_status("MiR_Mis_Queue") == 0)):
          sync()
        end
        $ 1125 "Set MiR_CMD_Clear_Q=Off"
        modbus_set_output_signal("MiR_CMD_Clear_Q", False)
      end
      $ 1126 "If MiR_Error_ID≠0"
      if (modbus_get_signal_status("MiR_Error_ID") != 0):
        $ 1127 "Set MiR_CMD_Clear_E=On"
        modbus_set_output_signal("MiR_CMD_Clear_E", True)
        $ 1128 "Wait MiR_Error_ID≟0"
        while (not(modbus_get_signal_status("MiR_Error_ID") == 0)):
          sync()
        end
        $ 1129 "Set MiR_CMD_Clear_E=Off"
        modbus_set_output_signal("MiR_CMD_Clear_E", False)
      end
      $ 1130 "Set O2T_Action=0"
      modbus_set_output_register("O2T_Action", 0)
      $ 1131 "Set O2T_Acknowledge=0"
      modbus_set_output_register("O2T_Acknowledge", 0)
      $ 1132 "Set O2T_Target_Pos=0"
      modbus_set_output_register("O2T_Target_Pos", 0)
      $ 1133 "Set O2T_Footprint=0"
      modbus_set_output_register("O2T_Footprint", 0)
      $ 1134 "Set O2T_ProtectOff=0"
      modbus_set_output_register("O2T_ProtectOff", 0)
      $ 1135 "Set O2T_Dock=0"
      modbus_set_output_register("O2T_Dock", 0)
      $ 1136 "AMR_Attemps≔0"
      global AMR_Attemps=0
      $ 1137 "AMR_PosTarget≔0"
      global AMR_PosTarget=0
      $ 1138 "AMR_Step≔0"
      global AMR_Step=0
      $ 1139 "AMR_AtTarget≔ False "
      global AMR_AtTarget=  False
      $ 1140 "If MiR_State≟4 or MiR_State≟3 or MiR_State≟10"
      if (modbus_get_signal_status("MiR_State") == 4  or  modbus_get_signal_status("MiR_State") == 3  or  modbus_get_signal_status("MiR_State") == 10):
        $ 1141 "AMR_Done≔ True "
        global AMR_Done=  True
      end
    elif (5 == switch_1):
      $ 1142 "Case 5"
      $ 1143 "starting"
      $ 1144 "If MiR_State≟4"
      if (modbus_get_signal_status("MiR_State") == 4):
        $ 1145 "Set MiR_CMD_Start=On"
        modbus_set_output_signal("MiR_CMD_Start", True)
        $ 1146 "Wait MiR_State≠4"
        while (not(modbus_get_signal_status("MiR_State") != 4)):
          sync()
        end
        $ 1147 "Set MiR_CMD_Start=Off"
        modbus_set_output_signal("MiR_CMD_Start", False)
        $ 1148 "AMR_Done≔ True "
        global AMR_Done=  True
      else:
        $ 1149 "ElseIf MiR_State≟10"
        if (modbus_get_signal_status("MiR_State") == 10):
          $ 1150 "'MiR in protective stop. Wait'"
          # 'MiR in protective stop. Wait'
          $ 1151 "AMR_Done≔ True "
          global AMR_Done=  True
        else:
          $ 1152 "ElseIf MiR_State≟3"
          if (modbus_get_signal_status("MiR_State") == 3):
            $ 1153 "AMR_Done≔ True "
            global AMR_Done=  True
          end
        end
      end
    elif (6 == switch_1):
      $ 1154 "Case 6"
      $ 1155 "execute"
      $ 1156 "AMR_AtTarget≔(AMR_PosActual≟AMR_PosTarget)"
      global AMR_AtTarget=(AMR_PosActual == AMR_PosTarget)
      $ 1157 "Switch AMR_Step"
      switch_2 = AMR_Step
      $ 1158 "Case 0"
      if (0 == switch_2):
        $ 1159 "If  not AMR_AtTarget"
        if (  not  AMR_AtTarget):
          $ 1160 "AMR_Step≔1"
          global AMR_Step=1
        else:
          $ 1161 "Else" "noBreak"
          $ 1162 "AMR_Done≔ True "
          global AMR_Done=  True
        end
      elif (1 == switch_2):
        $ 1163 "Case 1"
        $ 1164 "general Settings"
        $ 1165 "Set O2T_Acknowledge=0"
        modbus_set_output_register("O2T_Acknowledge", 0)
        $ 1166 "check for error"
        $ 1167 "If OBJ_Picked and MiR_State≟10"
        if (OBJ_Picked  and  modbus_get_signal_status("MiR_State") == 10):
          $ 1168 "Error"
          $ 1169 "set_error(ERROR_ROBOT_ARM_NOT_IN_HOME_POSE)"
          set_error(ERROR_ROBOT_ARM_NOT_IN_HOME_POSE)
          $ 1170 "Action≔0"
          global Action=0
        else:
          $ 1171 "ElseIf  not found_in_list(AMR_PosTarget, AMR_TargetList)"
          if (  not  found_in_list(AMR_PosTarget, AMR_TargetList)):
            $ 1172 "Error"
            $ 1173 "set_error(ERROR_UNKNOWN_POSE)"
            set_error(ERROR_UNKNOWN_POSE)
            $ 1174 "Action≔0"
            global Action=0
          end
        end
        $ 1175 "If MiR_State≟3"
        if (modbus_get_signal_status("MiR_State") == 3):
          $ 1176 "Set MiR_CMD_Start=Off"
          modbus_set_output_signal("MiR_CMD_Start", False)
          $ 1177 "Switch Action"
          switch_3 = Action
          $ 1178 "Case 51"
          if (51 == switch_3):
            $ 1179 "Charge"
            $ 1180 "'trigger the charging mission'"
            # 'trigger the charging mission'
            $ 1181 "'target pos is predefined'"
            # 'target pos is predefined'
            $ 1182 "Set O2T_Footprint=0"
            modbus_set_output_register("O2T_Footprint", 0)
            $ 1183 "Set O2T_Action=1"
            modbus_set_output_register("O2T_Action", 1)
            $ 1184 "If MiR_Mis_Queue≟0"
            if (modbus_get_signal_status("MiR_Mis_Queue") == 0):
              $ 1185 "Set O2T_Mis_Charge=On"
              modbus_set_output_signal("O2T_Mis_Charge", True)
              $ 1186 "Wait MiR_Mis_Queue≥1"
              while (not(modbus_get_signal_status("MiR_Mis_Queue") >= 1)):
                sync()
              end
              $ 1187 "Set O2T_Mis_Charge=Off"
              modbus_set_output_signal("O2T_Mis_Charge", False)
            end
          elif (52 == switch_3):
            $ 1188 "Case 52"
            $ 1189 "Navigate"
            $ 1190 "'trigger the standard missoin'"
            # 'trigger the standard missoin'
            $ 1191 "Set O2T_Footprint=AMR_FootprintID"
            modbus_set_output_register("O2T_Footprint", AMR_FootprintID)
            $ 1192 "Set O2T_Target_Pos=AMR_PosTarget"
            modbus_set_output_register("O2T_Target_Pos", AMR_PosTarget)
            $ 1193 "Set O2T_Action=2"
            modbus_set_output_register("O2T_Action", 2)
            $ 1194 "If MiR_Mis_Queue≟0"
            if (modbus_get_signal_status("MiR_Mis_Queue") == 0):
              $ 1195 "Set O2T_Mis_Main=On"
              modbus_set_output_signal("O2T_Mis_Main", True)
              $ 1196 "Wait MiR_Mis_Queue≥1"
              while (not(modbus_get_signal_status("MiR_Mis_Queue") >= 1)):
                sync()
              end
              $ 1197 "Set O2T_Mis_Main=Off"
              modbus_set_output_signal("O2T_Mis_Main", False)
            end
          end
        else:
          $ 1198 "ElseIf MiR_State≟4"
          if (modbus_get_signal_status("MiR_State") == 4):
            $ 1199 "Set MiR_CMD_Start=On"
            modbus_set_output_signal("MiR_CMD_Start", True)
          else:
            $ 1200 "ElseIf MiR_State≟5"
            if (modbus_get_signal_status("MiR_State") == 5):
              $ 1201 "AMR_Step≔2"
              global AMR_Step=2
            else:
              $ 1202 "ElseIf MiR_State≟10"
              if (modbus_get_signal_status("MiR_State") == 10):
                $ 1203 "'AMR still in safeguard stop'"
                # 'AMR still in safeguard stop'
              end
            end
          end
        end
      elif (2 == switch_2):
        $ 1204 "Case 2"
        $ 1205 "acknowledge handshake"
        $ 1206 "If T2O_Done≟1 and O2T_Acknowledge≟0"
        if (modbus_get_signal_status("T2O_Done") == 1  and  modbus_get_signal_status("O2T_Acknowledge") == 0):
          $ 1207 "Set O2T_Acknowledge=1"
          modbus_set_output_register("O2T_Acknowledge", 1)
        else:
          $ 1208 "ElseIf T2O_Done≟0 and O2T_Acknowledge≟1"
          if (modbus_get_signal_status("T2O_Done") == 0  and  modbus_get_signal_status("O2T_Acknowledge") == 1):
            $ 1209 "Set O2T_Acknowledge=0"
            modbus_set_output_register("O2T_Acknowledge", 0)
            $ 1210 "AMR_AtTarget≔(AMR_PosActual≟AMR_PosTarget)"
            global AMR_AtTarget=(AMR_PosActual == AMR_PosTarget)
            $ 1211 "AMR_Done≔ True "
            global AMR_Done=  True
          end
        end
      end
      $ 1212 "translate errors"
      $ 1213 "If AMR_Done"
      if (AMR_Done):
        $ 1214 "Switch T2O_Error_ID"
        switch_2 = modbus_get_signal_status("T2O_Error_ID")
        $ 1215 "Case 2003"
        if (2003 == switch_2):
          $ 1216 "error"
          $ 1217 "set_error(ERROR_NOT_DOCKED)"
          set_error(ERROR_NOT_DOCKED)
        elif (2007 == switch_2):
          $ 1218 "Case 2007"
          $ 1219 "error"
          $ 1220 "set_error(ERROR_NOT_REACHABLE_TARGET)"
          set_error(ERROR_NOT_REACHABLE_TARGET)
        elif (2008 == switch_2):
          $ 1221 "Case 2008"
          $ 1222 "error"
          $ 1223 "set_error(ERROR_CHARGING_NOT_STARTED)"
          set_error(ERROR_CHARGING_NOT_STARTED)
        end
      end
    elif (7 == switch_1):
      $ 1224 "Case 7"
      $ 1225 "completing"
      $ 1226 "If MiR_Mis_Queue>0"
      if (modbus_get_signal_status("MiR_Mis_Queue")>0):
        $ 1227 "Set MiR_CMD_Abort=On"
        modbus_set_output_signal("MiR_CMD_Abort", True)
        $ 1228 "Wait MiR_Mis_Queue≟0"
        while (not(modbus_get_signal_status("MiR_Mis_Queue") == 0)):
          sync()
        end
        $ 1229 "Set MiR_CMD_Abort=Off"
        modbus_set_output_signal("MiR_CMD_Abort", False)
      end
      $ 1230 "If MiR_State≟3 or MiR_State≟10"
      if (modbus_get_signal_status("MiR_State") == 3  or  modbus_get_signal_status("MiR_State") == 10):
        $ 1231 "AMR_Done≔ True "
        global AMR_Done=  True
      end
    elif (9 == switch_1):
      $ 1232 "Case 9"
      $ 1233 "holding"
      $ 1234 "Set MiR_CMD_Abort=On"
      modbus_set_output_signal("MiR_CMD_Abort", True)
      $ 1235 "If MiR_State≟3 or MiR_State≟10"
      if (modbus_get_signal_status("MiR_State") == 3  or  modbus_get_signal_status("MiR_State") == 10):
        $ 1236 "Set MiR_CMD_Abort=Off"
        modbus_set_output_signal("MiR_CMD_Abort", False)
        $ 1237 "AMR_Done≔ True "
        global AMR_Done=  True
      end
    elif (11 == switch_1):
      $ 1238 "Case 11"
      $ 1239 "unholding"
      $ 1240 "Set MiR_CMD_Start=On"
      modbus_set_output_signal("MiR_CMD_Start", True)
      $ 1241 "If MiR_State≠4"
      if (modbus_get_signal_status("MiR_State") != 4):
        $ 1242 "Set MiR_CMD_Start=Off"
        modbus_set_output_signal("MiR_CMD_Start", False)
        $ 1243 "AMR_Step≔0"
        global AMR_Step=0
        $ 1244 "AMR_Done≔ True "
        global AMR_Done=  True
      end
    elif (12 == switch_1):
      $ 1245 "Case 12"
      $ 1246 "suspending"
      $ 1247 "'none'"
      # 'none'
    elif (14 == switch_1):
      $ 1248 "Case 14"
      $ 1249 "unsuspending"
      $ 1250 "'none'"
      # 'none'
    elif (15 == switch_1):
      $ 1251 "Case 15"
      $ 1252 "aborting"
      $ 1253 "Set MiR_CMD_Abort=On"
      modbus_set_output_signal("MiR_CMD_Abort", True)
      $ 1254 "Wait MiR_State≟3"
      while (not(modbus_get_signal_status("MiR_State") == 3)):
        sync()
      end
      $ 1255 "Set MiR_CMD_Abort=Off"
      modbus_set_output_signal("MiR_CMD_Abort", False)
    elif (17 == switch_1):
      $ 1256 "Case 17"
      $ 1257 "clearing"
      $ 1258 "If MiR_Error_ID≠0"
      if (modbus_get_signal_status("MiR_Error_ID") != 0):
        $ 1259 "Set MiR_CMD_Clear_E=On"
        modbus_set_output_signal("MiR_CMD_Clear_E", True)
        $ 1260 "Wait MiR_Error_ID≟0"
        while (not(modbus_get_signal_status("MiR_Error_ID") == 0)):
          sync()
        end
        $ 1261 "Set MiR_CMD_Clear_E=Off"
        modbus_set_output_signal("MiR_CMD_Clear_E", False)
      end
      $ 1262 "If MiR_Error_ID≟0"
      if (modbus_get_signal_status("MiR_Error_ID") == 0):
        $ 1263 "AMR_Done≔ True "
        global AMR_Done=  True
      end
    end
    $ 1264 "'=========='"
    # '=========='
    $ 1265 "PostSettings"
    $ 1266 "AMR_Position≔struct(position_identifier=T2O_Current_Pos, x1=MiR_Position_X1, x2=MiR_Position_X2, y1=MiR_Position_Y1, y2=MiR_Position_Y2, theta1=MiR_Theta_1, theta2=MiR_Theta_2) "
    global AMR_Position=struct(position_identifier=modbus_get_signal_status("T2O_Current_Pos"), x1=modbus_get_signal_status("MiR_Position_X1"), x2=modbus_get_signal_status("MiR_Position_X2"), y1=modbus_get_signal_status("MiR_Position_Y1"), y2=modbus_get_signal_status("MiR_Position_Y2"), theta1=modbus_get_signal_status("MiR_Theta_1"), theta2=modbus_get_signal_status("MiR_Theta_2"))
  end
  def Sub_Action_V4():
    $ 1267 "Sub_Action_V4" "noBreak"
    $ 1268 "PreSettings"
    $ 1269 "init poses"
    $ 1270 "PSE_A≔p[0,0,0,0,0,0]"
    global PSE_A=p[0,0,0,0,0,0]
    $ 1271 "PSE_A_H≔p[0,0,0,0,0,0]"
    global PSE_A_H=p[0,0,0,0,0,0]
    $ 1272 "PSE_T≔p[0,0,0,0,0,0]"
    global PSE_T=p[0,0,0,0,0,0]
    $ 1273 "PSE_T_H≔p[0,0,0,0,0,0]"
    global PSE_T_H=p[0,0,0,0,0,0]
    $ 1274 "PSE_G≔p[0,0,0,0,0,0]"
    global PSE_G=p[0,0,0,0,0,0]
    $ 1275 "PSE_G_H≔p[0,0,0,0,0,0]"
    global PSE_G_H=p[0,0,0,0,0,0]
    $ 1276 "PSE_R≔p[0,0,0,0,0,0]"
    global PSE_R=p[0,0,0,0,0,0]
    $ 1277 "PSE_R_H≔p[0,0,0,0,0,0]"
    global PSE_R_H=p[0,0,0,0,0,0]
    $ 1278 "JNT_Q≔[0,0,0,0,0,0]"
    global JNT_Q=[0,0,0,0,0,0]
    $ 1279 "JNT_S≔[0,0,0,0,0,0]"
    global JNT_S=[0,0,0,0,0,0]
    $ 1280 "Gripping parameters"
    $ 1281 "OBJ = find_object_by_type(OBJs, OBJ_Type)"
    OBJ = find_object_by_type(OBJs, OBJ_Type)
    $ 1282 "GRP_Open_Pos≔OBJ.dimension.diameter * 1000 + 6"
    global GRP_Open_Pos=OBJ.dimension.diameter * 1000 + 6
    $ 1283 "GRP_Offset≔OBJ.gripper_offset"
    global GRP_Offset=OBJ.gripper_offset
    $ 1284 "rq_set_force_norm(50)"
     rq_set_force_norm (50)
    $ 1285 "rq_set_speed_norm(50)"
     rq_set_speed_norm (50)
    $ 1286 "Switch ITM_ID"
    switch_1 = ITM_ID
    $ 1287 "Case 1"
    if (1 == switch_1):
      $ 1288 "uML"
      $ 1289 "JIG2 = find_object_by_type(JIGs, JIG)"
      JIG2 = find_object_by_type(JIGs, JIG)
      $ 1290 "JIG_Offset≔JIG2.jig_offset"
      global JIG_Offset=JIG2.jig_offset
      $ 1291 "Switch JIG"
      switch_2 = JIG
      $ 1292 "Case 1"
      if (1 == switch_2):
        $ 1293 "3FG"
        $ 1294 "define poses"
        $ 1295 "FRM_Reference≔ULM_3FG"
        global FRM_Reference=ULM_3FG
        $ 1296 "JNT_Q≔JNT_HOME"
        global JNT_Q=JNT_HOME
        $ 1297 "PSE_T≔pose_trans(GRP_Offset, JIG_Offset)"
        global PSE_T= pose_trans (GRP_Offset, JIG_Offset)
        $ 1298 "PSE_A≔pose_trans(PSE_T, p[0,0,0.100,0,0,0])"
        global PSE_A= pose_trans (PSE_T, p[0,0,0.100,0,0,0])
        $ 1299 "PSE_R≔pose_add(PSE_T, p[0,0,0.100,0,0,0])"
        global PSE_R= pose_add (PSE_T, p[0,0,0.100,0,0,0])
      elif (2 == switch_2):
        $ 1300 "Case 2"
        $ 1301 "Input"
        $ 1302 "'CHANGE THE REFERENCE TO THE FRAME TO MOVE IN'"
        # 'CHANGE THE REFERENCE TO THE FRAME TO MOVE IN'
        $ 1303 "define poses"
        $ 1304 "FRM_Reference≔ULM_Input"
        global FRM_Reference=ULM_Input
        $ 1305 "PSE_T≔pose_trans(pose_trans(get_pattern_pos_rectangle(OBJ_Nbr, 'X', [10,5], patternsize=[0.181,0.081]), GRP_Offset), JIG_Offset)"
        global PSE_T= pose_trans ( pose_trans (get_pattern_pos_rectangle(OBJ_Nbr, "X", [10,5], patternsize=[0.181,0.081]), GRP_Offset), JIG_Offset)
        $ 1306 "If Action≟1"
        if (Action == 1):
          $ 1307 "PSE_R≔pose_add(PSE_T, p[0,0,0.200,0,0,0])"
          global PSE_R= pose_add (PSE_T, p[0,0,0.200,0,0,0])
          $ 1308 "PSE_A≔pose_add(PSE_T, p[0,0,0.100,0,0,0])"
          global PSE_A= pose_add (PSE_T, p[0,0,0.100,0,0,0])
        else:
          $ 1309 "ElseIf Action≟2"
          if (Action == 2):
            $ 1310 "PSE_R≔pose_add(PSE_T, p[0,0,0.100,0,0,0])"
            global PSE_R= pose_add (PSE_T, p[0,0,0.100,0,0,0])
            $ 1311 "PSE_A≔pose_add(PSE_T, p[0,0,0.200,0,0,0])"
            global PSE_A= pose_add (PSE_T, p[0,0,0.200,0,0,0])
          end
        end
      elif (3 == switch_2):
        $ 1312 "Case 3"
        $ 1313 "Output"
        $ 1314 "'CHANGE THE REFERENCE TO THE FRAME TO MOVE IN'"
        # 'CHANGE THE REFERENCE TO THE FRAME TO MOVE IN'
        $ 1315 "define poses"
        $ 1316 "FRM_Reference≔ULM_Output"
        global FRM_Reference=ULM_Output
        $ 1317 "PSE_T≔pose_trans(pose_trans(get_pattern_pos_rectangle(OBJ_Nbr, 'X', [10,5], patternsize=[0.181,0.081]), GRP_Offset), JIG_Offset)"
        global PSE_T= pose_trans ( pose_trans (get_pattern_pos_rectangle(OBJ_Nbr, "X", [10,5], patternsize=[0.181,0.081]), GRP_Offset), JIG_Offset)
        $ 1319 "If Action≟1"
        if (Action == 1):
          $ 1320 "PSE_R≔pose_add(PSE_T, p[0,0,0.200,0,0,0])"
          global PSE_R= pose_add (PSE_T, p[0,0,0.200,0,0,0])
          $ 1321 "PSE_A≔pose_add(PSE_T, p[0,0,0.100,0,0,0])"
          global PSE_A= pose_add (PSE_T, p[0,0,0.100,0,0,0])
        else:
          $ 1322 "ElseIf Action≟2"
          if (Action == 2):
            $ 1323 "PSE_R≔pose_add(PSE_T, p[0,0,0.100,0,0,0])"
            global PSE_R= pose_add (PSE_T, p[0,0,0.100,0,0,0])
            $ 1324 "PSE_A≔pose_add(PSE_T, p[0,0,0.200,0,0,0])"
            global PSE_A= pose_add (PSE_T, p[0,0,0.200,0,0,0])
          end
        end
      elif (4 == switch_2):
        $ 1325 "Case 4"
        $ 1326 "jig centrifuge racks"
        $ 1327 "define poses"
        $ 1328 "FRM_Reference≔ULM_Cent_Racks"
        global FRM_Reference=ULM_Cent_Racks
        $ 1329 "PSE_T≔get_pattern_pos_rectangle(JIG_Slot, 'X', [4,1], patternsize=[0.291,0])"
        global PSE_T=get_pattern_pos_rectangle(JIG_Slot, "X", [4,1], patternsize=[0.291,0])
        $ 1330 "If OBJ_Nbr≠0"
        if (OBJ_Nbr != 0):
          $ 1331 "PSE_T≔pose_trans(pose_trans(PSE_T, get_pattern_pos_rectangle(OBJ_Nbr, 'X', [3,3], patternsize=[0.060,0.060])),p[-0.030, -0.030,0,0,0,3.927])"
          global PSE_T= pose_trans ( pose_trans (PSE_T, get_pattern_pos_rectangle(OBJ_Nbr, "X", [3,3], patternsize=[0.060,0.060])),p[-0.030, -0.030,0,0,0,3.927])
        end
        $ 1332 "PSE_T≔pose_trans(PSE_T, GRP_Offset)"
        global PSE_T= pose_trans (PSE_T, GRP_Offset)
        $ 1333 "If Action≟1"
        if (Action == 1):
          $ 1334 "PSE_R≔pose_add(PSE_T, p[0,0,0.200,0,0,0])"
          global PSE_R= pose_add (PSE_T, p[0,0,0.200,0,0,0])
          $ 1335 "PSE_A≔pose_add(PSE_T, p[0,0,0.100,0,0,0])"
          global PSE_A= pose_add (PSE_T, p[0,0,0.100,0,0,0])
        else:
          $ 1336 "ElseIf Action≟2"
          if (Action == 2):
            $ 1337 "PSE_R≔pose_add(PSE_T, p[0,0,0.100,0,0,0])"
            global PSE_R= pose_add (PSE_T, p[0,0,0.100,0,0,0])
            $ 1338 "PSE_A≔pose_add(PSE_T, p[0,0,0.200,0,0,0])"
            global PSE_A= pose_add (PSE_T, p[0,0,0.200,0,0,0])
          end
        end
      elif (6 == switch_2):
        $ 1339 "Case 6"
        $ 1340 "Caps bin"
        $ 1341 "define poses"
        $ 1342 "'Drop cap'"
        # 'Drop cap'
        $ 1343 "FRM_Reference=ULM_Cap_Bin"
        FRM_Reference=ULM_Cap_Bin
        $ 1344 "PSE_T≔pose_RPY2RotVec(p[0,0,0,0,0,0])"
        global PSE_T=pose_RPY2RotVec(p[0,0,0,0,0,0])
        $ 1345 "PSE_T_H≔pose_add(PSE_T, p[0,0,-0.011,0,0,0])"
        global PSE_T_H= pose_add (PSE_T, p[0,0,-0.011,0,0,0])
        $ 1346 "PSE_A≔pose_trans(PSE_T, p[0,0,0.1,0,0,0])"
        global PSE_A= pose_trans (PSE_T, p[0,0,0.1,0,0,0])
        $ 1347 "PSE_R_H≔pose_add(PSE_T, p[0,0,0.100,0,0,0])"
        global PSE_R_H= pose_add (PSE_T, p[0,0,0.100,0,0,0])
        $ 1348 "PSE_R≔pose_add(PSE_T, p[0,0,0.100,0,0,0])"
        global PSE_R= pose_add (PSE_T, p[0,0,0.100,0,0,0])
      elif (7 == switch_2):
        $ 1349 "Case 7"
        $ 1350 "Sarstedt"
        $ 1351 "'CHANGE THE REFERENCE TO THE FRAME TO MOVE IN'"
        # 'CHANGE THE REFERENCE TO THE FRAME TO MOVE IN'
        $ 1357 "If TASK.ID≟10"
        if (TASK.ID == 10):
          $ 1358 "Frame & Position Params"
          $ 1360 "FRM_Reference = CAM_LM_SSRack"
          FRM_Reference = CAM_LM_SSRack
          $ 1365 "PSE_T≔uLM_SS_PickPlc"
          global PSE_T=uLM_SS_PickPlc
          $ 1366 "PSE_A≔pose_trans(PSE_T, p[0,0,0.1,0,0,0])"
          global PSE_A= pose_trans (PSE_T, p[0,0,0.1,0,0,0])
          $ 1367 "PSE_R≔pose_add(PSE_T, p[0,0,0.1,0,0,0])"
          global PSE_R= pose_add (PSE_T, p[0,0,0.1,0,0,0])
        else:
          $ 1368 "ElseIf TASK.ID≟11"
          if (TASK.ID == 11):
            $ 1369 "FRM_Reference = ULM_SS_Jig"
            FRM_Reference = ULM_SS_Jig
            $ 1370 "PSE_T≔pose_RPY2RotVec(p[0,0,0,0,0,0])"
            global PSE_T=pose_RPY2RotVec(p[0,0,0,0,0,0])
            $ 1371 "PSE_T≔pose_trans(PSE_T, GRP_Offset)"
            global PSE_T=pose_trans(PSE_T, GRP_Offset)
            $ 1372 "PSE_A≔pose_trans(PSE_T, p[0,0,0.1,0,0,0])"
            global PSE_A= pose_trans (PSE_T, p[0,0,0.1,0,0,0])
            $ 1373 "PSE_R≔pose_add(PSE_T, p[0,0,0.2,0,0,0])"
            global PSE_R= pose_add (PSE_T, p[0,0,0.2,0,0,0])
          end
        end
      elif (8 == switch_2):
        $ 1374 "Case 8"
        $ 1375 "NoK"
        $ 1376 "define poses"
        $ 1377 "'NoK'"
        # 'NoK'
        $ 1378 "FRM_Reference=ULM_NoK"
        FRM_Reference=ULM_NoK
        $ 1379 "PSE_T≔pose_RPY2RotVec(p[0,0,0,0,0,0])"
        global PSE_T=pose_RPY2RotVec(p[0,0,0,0,0,0])
        $ 1380 "PSE_A≔pose_trans(PSE_T, p[0,0,0.1,0,0,0])"
        global PSE_A= pose_trans (PSE_T, p[0,0,0.1,0,0,0])
        $ 1381 "PSE_R≔pose_add(PSE_T, p[0,0,0.100,0,0,0])"
        global PSE_R= pose_add (PSE_T, p[0,0,0.100,0,0,0])
      elif (9 == switch_2):
        $ 1382 "Case 9"
        $ 1383 "Pick_bott_jig"
        $ 1384 "define poses"
        $ 1385 "'NoK'"
        # 'NoK'
        $ 1386 "FRM_Reference=ULM_bottle_pick_const"
        FRM_Reference=p[0.08175869478771049,-0.47602162643540935,0.09,0.00141829700319658,-0.0027789445191063835,0.07763675748118615]
        $ 1387 "PSE_T≔pose_RPY2RotVec(p[0,0,0,0,0,0])"
        global PSE_T=pose_RPY2RotVec(p[0,0,0,0,0,0])
        $ 1388 "PSE_A≔pose_trans(PSE_T, p[0,0,0.1,0,0,0])"
        global PSE_A= pose_trans (PSE_T, p[0,0,0.1,0,0,0])
        $ 1389 "PSE_R≔pose_add(PSE_T, p[0,0,0.100,0,0,0])"
        global PSE_R= pose_add (PSE_T, p[0,0,0.100,0,0,0])
      elif (10 == switch_2):
        $ 1390 "Case 10"
        $ 1391 "Place_bott_jig"
        $ 1392 "define poses"
        $ 1393 "'NoK'"
        # 'NoK'
        $ 1394 "FRM_Reference=ULM_bottle_plac_const"
        FRM_Reference=p[-0.09502738395762109,-0.5154087721098056,0.095,0.0014590126708889871,-0.0028280855286173575,0.07763149296298452]
        $ 1395 "PSE_T≔pose_RPY2RotVec(p[0,0,0,0,0,0])"
        global PSE_T=pose_RPY2RotVec(p[0,0,0,0,0,0])
        $ 1396 "PSE_A≔pose_trans(PSE_T, p[0,0,0.1,0,0,0])"
        global PSE_A= pose_trans (PSE_T, p[0,0,0.1,0,0,0])
        $ 1397 "PSE_R≔pose_add(PSE_T, p[0,0,0.100,0,0,0])"
        global PSE_R= pose_add (PSE_T, p[0,0,0.100,0,0,0])
      elif (11 == switch_2):
        $ 1398 "Case 11"
        $ 1399 "Place_bott_jig"
        $ 1400 "define poses"
        $ 1401 "'NoK'"
        # 'NoK'
        $ 1402 "FRM_Reference=shake"
        FRM_Reference=shake
        $ 1403 "PSE_T≔pose_RPY2RotVec(p[0,0,0,0,0,0])"
        global PSE_T=pose_RPY2RotVec(p[0,0,0,0,0,0])
        $ 1404 "PSE_A≔pose_trans(PSE_T, p[0,0,0,0,0,0])"
        global PSE_A= pose_trans (PSE_T, p[0,0,0,0,0,0])
        $ 1405 "PSE_R≔pose_add(PSE_T, p[0,0,0,0,0,0])"
        global PSE_R= pose_add (PSE_T, p[0,0,0,0,0,0])
      elif (12 == switch_2):
        $ 1406 "Case 12"
        $ 1407 "Pick_Vial_jig"
        $ 1408 "define poses"
        $ 1409 "'NoK'"
        # 'NoK'
        $ 1410 "FRM_Reference=shake"
        FRM_Reference=shake
        $ 1411 "PSE_T≔pose_RPY2RotVec(p[0,0,0,0,0,0])"
        global PSE_T=pose_RPY2RotVec(p[0,0,0,0,0,0])
        $ 1412 "PSE_A≔pose_trans(PSE_T, p[0,0,0,0,0,0])"
        global PSE_A= pose_trans (PSE_T, p[0,0,0,0,0,0])
        $ 1413 "PSE_R≔pose_add(PSE_T, p[0,0,0,0,0,0])"
        global PSE_R= pose_add (PSE_T, p[0,0,0,0,0,0])
      end
    elif (2 == switch_1):
      $ 1414 "Case 2"
      $ 1415 "Centrifuge"
      $ 1416 "'CHANGE THE REFERENCE TO THE FRAME TO MOVE IN'"
      # 'CHANGE THE REFERENCE TO THE FRAME TO MOVE IN'
      $ 1417 "define poses"
      $ 1418 "FRM_Reference≔FRM_Centrifuge"
      global FRM_Reference=FRM_Centrifuge
      $ 1419 "PSE_T≔GRP_Offset"
      global PSE_T=GRP_Offset
      $ 1420 "If Action≟8"
      if (Action == 8):
        $ 1421 "PSE_R≔pose_add(PSE_T, p[0,0,0.250,0,0,0])"
        global PSE_R= pose_add (PSE_T, p[0,0,0.250,0,0,0])
        $ 1422 "PSE_A≔pose_add(PSE_T, p[0,0,0.150,0,0,0])"
        global PSE_A= pose_add (PSE_T, p[0,0,0.150,0,0,0])
      else:
        $ 1423 "ElseIf Action≟7"
        if (Action == 7):
          $ 1424 "PSE_R≔pose_add(PSE_T, p[0,0,0.150,0,0,0])"
          global PSE_R= pose_add (PSE_T, p[0,0,0.150,0,0,0])
          $ 1425 "PSE_A≔pose_add(PSE_T, p[0,0,0.250,0,0,0])"
          global PSE_A= pose_add (PSE_T, p[0,0,0.250,0,0,0])
        end
      end
    elif (3 == switch_1):
      $ 1426 "Case 3"
      $ 1427 "Output"
      $ 1428 "'CHANGE THE REFERENCE TO THE FRAME TO MOVE IN'"
      # 'CHANGE THE REFERENCE TO THE FRAME TO MOVE IN'
      $ 1429 "define poses"
      $ 1430 "FRM_Reference≔Base_const"
      global FRM_Reference=p[0.0,0.0,0.0,0.0,0.0,0.0]
      $ 1431 "PSE_T≔p[0,0,0,0,0,0]"
      global PSE_T=p[0,0,0,0,0,0]
      $ 1432 "PSE_A≔pose_add(PSE_T, p[0,0,0.150,0,0,0])"
      global PSE_A= pose_add (PSE_T, p[0,0,0.150,0,0,0])
      $ 1433 "PSE_R≔pose_add(PSE_T, p[0,0,0.100,0,0,0])"
      global PSE_R= pose_add (PSE_T, p[0,0,0.100,0,0,0])
    elif (5 == switch_1):
      $ 1434 "Case 5"
      $ 1435 "Sarstedt Pickup Table"
      $ 1436 "'CHANGE THE REFERENCE TO THE FRAME TO MOVE IN'"
      # 'CHANGE THE REFERENCE TO THE FRAME TO MOVE IN'
      $ 1437 "Switch JIG"
      switch_2 = JIG
      $ 1438 "Case 7"
      if (7 == switch_2):
        $ 1451 "Sarstedt"
        $ 1452 "'CHANGE THE REFERENCE TO THE FRAME TO MOVE IN'"
        # 'CHANGE THE REFERENCE TO THE FRAME TO MOVE IN'
        $ 1458 "If TASK.ID≟10"
        if (TASK.ID == 10):
          $ 1459 "Frame & Position Params"
          $ 1460 "FRM_Reference = CAM_LM_SSRack"
          FRM_Reference = CAM_LM_SSRack
          $ 1461 "PSE_T≔uLM_SS_PickPlc"
          global PSE_T=uLM_SS_PickPlc
          $ 1462 "PSE_A≔pose_trans(PSE_T, p[0,0,0.1,0,0,0])"
          global PSE_A= pose_trans (PSE_T, p[0,0,0.1,0,0,0])
          $ 1463 "PSE_R≔pose_add(PSE_T, p[0,0,0.1,0,0,0])"
          global PSE_R= pose_add (PSE_T, p[0,0,0.1,0,0,0])
        end
      end
    elif (13 == switch_1):
      $ 1470 "Case 13"
      $ 1471 "Sarstedt Pickup Table"
      $ 1472 "'CHANGE THE REFERENCE TO THE FRAME TO MOVE IN'"
      # 'CHANGE THE REFERENCE TO THE FRAME TO MOVE IN'
      $ 1473 "Switch JIG"
      switch_2 = JIG
      $ 1474 "Case 7"
      if (7 == switch_2):
        $ 1487 "Bottle"
        $ 1488 "'CHANGE THE REFERENCE TO THE FRAME TO MOVE IN'"
        # 'CHANGE THE REFERENCE TO THE FRAME TO MOVE IN'
        $ 1494 "If TASK.ID≟43"
        if (TASK.ID == 43):
          $ 1495 "Frame & Position Params"
          $ 1496 "FRM_Reference = CAM_LM_Bott"
          FRM_Reference = CAM_LM_Bott
          $ 1497 "PSE_T≔uLM_SS_PickPlc"
          global PSE_T=uLM_SS_PickPlc
          $ 1498 "PSE_A≔pose_trans(PSE_T, p[0,0,0.1,0,0,0])"
          global PSE_A= pose_trans (PSE_T, p[0,0,0.1,0,0,0])
          $ 1499 "PSE_R≔pose_add(PSE_T, p[0,0,0.1,0,0,0])"
          global PSE_R= pose_add (PSE_T, p[0,0,0.1,0,0,0])
        end
      end
    end
    $ 1506 "Additional check"
    $ 1507 "If  not is_reachable(FRM_Reference,[PSE_A,PSE_A_H,PSE_T,PSE_T_H,PSE_R,PSE_R_H])"
    if (  not  is_reachable(FRM_Reference,[PSE_A,PSE_A_H,PSE_T,PSE_T_H,PSE_R,PSE_R_H])):
      $ 1508 "Error"
      $ 1509 "set_error(ERROR_POSE_NOT_REACHABLE)"
      set_error(ERROR_POSE_NOT_REACHABLE)
      $ 1510 "Action≔0"
      global Action=0
    end
    $ 1511 "'=========='"
    # '=========='
    $ 1512 "Switch Action"
    switch_1 = Action
    $ 1513 "Case 1"
    if (1 == switch_1):
      $ 1514 "Pick"
      $ 1515 "Action_Info≔'pick object'"
      global Action_Info="pick object"
      $ 1516 "do_transition(pose_trans(FRM_Reference, PSE_T), keep_rxry=OBJ_Picked)"
      do_transition( pose_trans (FRM_Reference, PSE_T), keep_rxry=OBJ_Picked)
      $ 1517 "EOAT"
      $ 1518 "If  not OBJ_Picked"
      if (  not  OBJ_Picked):
        $ 1519 "rq_move_and_wait_mm(GRP_Open_Pos)"
         rq_move_and_wait_mm (GRP_Open_Pos)
      end
      $ 1520 "If PSE_A_H≠PSE_Z"
      if (PSE_A_H != PSE_Z):
        $ 1521 "If JNT_Q≠JNT_Z"
        if (JNT_Q != JNT_Z):
          $ 1522 "movej(get_inverse_kin(pose_trans(FRM_Reference, PSE_A_H), qnear=JNT_Q), r=0.050)"
          movej(get_inverse_kin( pose_trans (FRM_Reference, PSE_A_H), qnear=JNT_Q), r=0.050)
        else:
          $ 1523 "Else" "noBreak"
          $ 1524 "movej(pose_trans(FRM_Reference, PSE_A_H), r=0.050)"
          movej( pose_trans (FRM_Reference, PSE_A_H), r=0.050)
        end
      end
      $ 1525 "If PSE_A≠PSE_Z"
      if (PSE_A != PSE_Z):
        $ 1526 "If JNT_Q≠JNT_Z"
        if (JNT_Q != JNT_Z):
          $ 1527 "movej(get_inverse_kin(pose_trans(FRM_Reference, PSE_A), qnear=JNT_Q), r=0.020)"
          movej(get_inverse_kin( pose_trans (FRM_Reference, PSE_A), qnear=JNT_Q), r=0.020)
        else:
          $ 1528 "Else" "noBreak"
          $ 1529 "movej(pose_trans(FRM_Reference, PSE_A), r=0.020)"
          movej( pose_trans (FRM_Reference, PSE_A), r=0.020)
        end
      end
      $ 1530 "MoveL"
      $ 1531 "If PSE_T_H≠PSE_Z"
      if (PSE_T_H != PSE_Z):
        $ 1532 "PSE_T_H" "breakAfter"
        movel(pose_trans(FRM_Reference, PSE_T_H), a=0.5, v=0.4, r=0.01)
      end
      $ 1533 "PSE_T" "breakAfter"
      movel(pose_trans(FRM_Reference, PSE_T), a=0.08, v=0.12)
      $ 1534 "EOAT"
      $ 1535 "rq_set_force_norm(50)"
       rq_set_force_norm (50)
      $ 1536 "rq_close_and_wait()"
       rq_close_and_wait ()
      $ 1537 "OBJ_Picked≔rq_is_object_detected()"
      global OBJ_Picked= rq_is_object_detected ()
      $ 1538 "If  not OBJ_Picked"
      if (  not  OBJ_Picked):
        $ 1539 "set_error(ERROR_NO_OBJECT_TO_PICK)"
        set_error(ERROR_NO_OBJECT_TO_PICK)
      end
      $ 1540 "EXTT"
      $ 1541 "Switch JIG"
      switch_2 = JIG
      $ 1542 "Case 1"
      if (1 == switch_2):
        $ 1543 "3FG"
        $ 1544 "If OBJ_Picked"
        if (OBJ_Picked):
          $ 1545 "Set GRP_3F_Open=On"
          set_standard_digital_out(5, True)
        end
      end
      $ 1546 "If PSE_R_H≠PSE_Z"
      if (PSE_R_H != PSE_Z):
        $ 1547 "PSE_R" "breakAfter"
        movel(pose_trans(FRM_Reference, PSE_R), a=0.5, v=0.4, r=0.01)
        $ 1548 "PSE_R_H" "breakAfter"
        movel(pose_trans(FRM_Reference, PSE_R_H), a=0.5, v=0.4)
      else:
        $ 1549 "Else" "noBreak"
        $ 1550 "PSE_R" "breakAfter"
        movel(pose_trans(FRM_Reference, PSE_R), a=0.5, v=0.4)
      end
    elif (2 == switch_1):
      $ 1551 "Case 2"
      $ 1552 "Place"
      $ 1553 "Action_Info≔'place object'"
      global Action_Info="place object"
      $ 1554 "do_transition(pose_trans(FRM_Reference, PSE_T), keep_rxry=OBJ_Picked)"
      do_transition( pose_trans (FRM_Reference, PSE_T), keep_rxry=OBJ_Picked)
      $ 1555 "EXTT"
      $ 1556 "Switch JIG"
      switch_2 = JIG
      $ 1557 "Case 1"
      if (1 == switch_2):
        $ 1558 "3FG"
        $ 1559 "If OBJ_Picked"
        if (OBJ_Picked):
          $ 1560 "Set GRP_3F_Open=On"
          set_standard_digital_out(5, True)
        end
      end
      $ 1561 "If PSE_A_H≠PSE_Z"
      if (PSE_A_H != PSE_Z):
        $ 1562 "If JNT_Q≠JNT_Z"
        if (JNT_Q != JNT_Z):
          $ 1563 "movej(get_inverse_kin(pose_trans(FRM_Reference, PSE_A_H), qnear=JNT_Q), r=0.050)"
          movej(get_inverse_kin( pose_trans (FRM_Reference, PSE_A_H), qnear=JNT_Q), r=0.050)
        else:
          $ 1564 "Else" "noBreak"
          $ 1565 "movej(pose_trans(FRM_Reference, PSE_A_H), r=0.050)"
          movej( pose_trans (FRM_Reference, PSE_A_H), r=0.050)
        end
      end
      $ 1566 "If PSE_A≠PSE_Z"
      if (PSE_A != PSE_Z):
        $ 1567 "If JNT_Q≠JNT_Z"
        if (JNT_Q != JNT_Z):
          $ 1568 "movej(get_inverse_kin(pose_trans(FRM_Reference, PSE_A), qnear=JNT_Q), r=0.020)"
          movej(get_inverse_kin( pose_trans (FRM_Reference, PSE_A), qnear=JNT_Q), r=0.020)
        else:
          $ 1569 "Else" "noBreak"
          $ 1570 "movej(pose_trans(FRM_Reference, PSE_A), r=0.020)"
          movej( pose_trans (FRM_Reference, PSE_A), r=0.020)
        end
      end
      $ 1571 "MoveL"
      $ 1572 "If PSE_T_H≠PSE_Z"
      if (PSE_T_H != PSE_Z):
        $ 1573 "PSE_T_H" "breakAfter"
        movel(pose_trans(FRM_Reference, PSE_T_H), a=0.5, v=0.4, r=0.01)
      end
      $ 1574 "PSE_T" "breakAfter"
      global move_thread_flag_1574=0
      thread move_thread_1574():
        enter_critical
        move_thread_flag_1574 = 1
        movel(pose_trans(FRM_Reference, PSE_T), a=0.05, v=0.09)
        move_thread_flag_1574 = 2
        exit_critical
      end
      move_thread_flag_1574 = 0
      move_thread_han_1574 = run move_thread_1574()
      while (True):
        local targetTcpDirection=get_target_tcp_speed()
        local stepsToRetract=tool_contact(direction=targetTcpDirection)
        if (stepsToRetract > 0):
          kill move_thread_han_1574
          stopl(0.5)
          $ 1575 "Until (tool_contact_detection)"
          break
        end
        sleep(1.0E-10)
        if (move_thread_flag_1574 > 1):
          join move_thread_han_1574
          break
        end
        sync()
      end
      $ 1576 "Force"
      sleep(0.02)
      zero_ftsensor()
      force_mode(FRM_Reference, [1, 1, 1, 0, 0, 0], [0.0, 0.0, 0.0, 0.0, 0.0, 0.0], 2, [0.1, 0.1, 0.01, 0.3490658503988659, 0.3490658503988659, 0.3490658503988659])
      $ 1577 "PSE_T" "noBreak"
      movel(pose_trans(FRM_Reference, PSE_T), a=0.04, v=0.07)
      end_force_mode()
      stopl(5.0)
      $ 1578 "EXTT"
      $ 1579 "Switch JIG"
      switch_2 = JIG
      $ 1580 "Case 1"
      if (1 == switch_2):
        $ 1581 "3FG"
        $ 1582 "If OBJ_Picked"
        if (OBJ_Picked):
          $ 1583 "Set GRP_3F_Open=Off"
          set_standard_digital_out(5, False)
          $ 1584 "Wait: 0.2"
          sleep(0.2)
        end
      end
      $ 1585 "EOAT"
      $ 1586 "rq_move_and_wait_mm(GRP_Open_Pos)"
       rq_move_and_wait_mm (GRP_Open_Pos)
      $ 1587 "OBJ_Picked≔rq_is_object_detected()"
      global OBJ_Picked= rq_is_object_detected ()
      $ 1588 "If PSE_R_H≠PSE_Z"
      if (PSE_R_H != PSE_Z):
        $ 1589 "PSE_R" "breakAfter"
        movel(pose_trans(FRM_Reference, PSE_R), a=0.5, v=0.4, r=0.01)
        $ 1590 "PSE_R_H" "breakAfter"
        movel(pose_trans(FRM_Reference, PSE_R_H), a=0.5, v=0.4)
      else:
        $ 1591 "Else" "noBreak"
        $ 1592 "PSE_R" "breakAfter"
        movel(pose_trans(FRM_Reference, PSE_R), a=0.5, v=0.4)
      end
    elif (3 == switch_1):
      $ 1593 "Case 3"
      $ 1594 "Push"
      $ 1595 "Action_Info≔'push'"
      global Action_Info="push"
    elif (4 == switch_1):
      $ 1596 "Case 4"
      $ 1597 "Pull"
      $ 1598 "Action_Info≔'pull'"
      global Action_Info="pull"
    elif (6 == switch_1):
      $ 1601 "Case 6"
      $ 1602 "Drop the cap"
      $ 1603 "If JNT_A≠[0,0,0,0,0,0]"
      if (JNT_A != [0,0,0,0,0,0]):
        $ 1604 "MoveJ"
        $ 1605 "JNT_A" "breakAfter"
        movej(JNT_A, a=1.3962634015954636, v=1.7453292519943295, r=0.02)
      else:
        $ 1606 "Else" "noBreak"
        $ 1607 "MoveJ"
        $ 1608 "PSE_A" "breakAfter"
        movej(pose_trans(FRM_Reference, PSE_A), a=1.3962634015954636, v=1.7453292519943295, r=0.02)
      end
      $ 1609 "MoveL"
      $ 1610 "PSE_T" "breakAfter"
      movel(pose_trans(FRM_Reference, PSE_T), a=0.05, v=0.09)
      $ 1611 "'ADD OPEN GRIPPER'"
      # 'ADD OPEN GRIPPER'
      # begin: URCap Program Node
      #   Source: Robotiq_Grippers, 1.8.4.4844, Robotiq Inc.
      #   Type: Gripper
      $ 1612 "Gripper Move10mm (1)"
      if not(gripper_connected[0]):
        popup("Gripper 1 must be connected to run this program.", "No connection", False, True, True)
      end
      if not(rq_is_gripper_activated("1")):
        popup("Gripper 1 is not activated. Go to Installation tab > Gripper to activate it and run the program again.", "Not activated", False, True, True)
      end
      rq_set_pos_spd_for(201, 0, 28, "1")
      rq_wait_pos_spe_for_request(201, 0, 28, "1")
      rq_go_to("1")
      rq_wait("1")
      # end: URCap Program Node
      $ 1613 "PSE_T_H" "breakAfter"
      movel(pose_trans(FRM_Reference, PSE_T_H), a=0.05, v=0.09)
      # begin: URCap Program Node
      #   Source: Robotiq_Grippers, 1.8.4.4844, Robotiq Inc.
      #   Type: Gripper
      $ 1614 "Gripper Move40mm (1)"
      if not(gripper_connected[0]):
        popup("Gripper 1 must be connected to run this program.", "No connection", False, True, True)
      end
      if not(rq_is_gripper_activated("1")):
        popup("Gripper 1 is not activated. Go to Installation tab > Gripper to activate it and run the program again.", "Not activated", False, True, True)
      end
      rq_set_pos_spd_for(63, 0, 28, "1")
      rq_wait_pos_spe_for_request(63, 0, 28, "1")
      rq_go_to("1")
      rq_wait("1")
      # end: URCap Program Node
      $ 1615 "PSE_R" "breakAfter"
      movel(pose_trans(FRM_Reference, PSE_R), a=0.5, v=0.4)
    elif (7 == switch_1):
      $ 1616 "Case 7"
      $ 1617 "Load"
      $ 1618 "Action_Info≔'load object'"
      global Action_Info="load object"
      $ 1619 "do_transition(pose_trans(FRM_Reference, PSE_T), keep_rxry=OBJ_Picked)"
      do_transition( pose_trans (FRM_Reference, PSE_T), keep_rxry=OBJ_Picked)
      $ 1620 "If PSE_A_H≠PSE_Z"
      if (PSE_A_H != PSE_Z):
        $ 1621 "If JNT_Q≠JNT_Z"
        if (JNT_Q != JNT_Z):
          $ 1622 "movej(get_inverse_kin(pose_trans(FRM_Reference, PSE_A_H), qnear=JNT_Q), r=0.050)"
          movej(get_inverse_kin( pose_trans (FRM_Reference, PSE_A_H), qnear=JNT_Q), r=0.050)
        else:
          $ 1623 "Else" "noBreak"
          $ 1624 "movej(pose_trans(FRM_Reference, PSE_A_H), r=0.050)"
          movej( pose_trans (FRM_Reference, PSE_A_H), r=0.050)
        end
      end
      $ 1625 "If PSE_A≠PSE_Z"
      if (PSE_A != PSE_Z):
        $ 1626 "If JNT_Q≠JNT_Z"
        if (JNT_Q != JNT_Z):
          $ 1627 "movej(get_inverse_kin(pose_trans(FRM_Reference, PSE_A), qnear=JNT_Q), r=0.020)"
          movej(get_inverse_kin( pose_trans (FRM_Reference, PSE_A), qnear=JNT_Q), r=0.020)
        else:
          $ 1628 "Else" "noBreak"
          $ 1629 "movej(pose_trans(FRM_Reference, PSE_A), r=0.020)"
          movej( pose_trans (FRM_Reference, PSE_A), r=0.020)
        end
      end
      $ 1630 "MoveL"
      $ 1631 "If PSE_T_H≠PSE_Z"
      if (PSE_T_H != PSE_Z):
        $ 1632 "PSE_T_H" "breakAfter"
        movel(pose_trans(FRM_Reference, PSE_T_H), a=0.5, v=0.4, r=0.01)
      end
      $ 1633 "PSE_T" "breakAfter"
      global move_thread_flag_1633=0
      thread move_thread_1633():
        enter_critical
        move_thread_flag_1633 = 1
        movel(pose_trans(FRM_Reference, PSE_T), a=0.05, v=0.09)
        move_thread_flag_1633 = 2
        exit_critical
      end
      move_thread_flag_1633 = 0
      move_thread_han_1633 = run move_thread_1633()
      while (True):
        local targetTcpDirection=get_target_tcp_speed()
        local stepsToRetract=tool_contact(direction=targetTcpDirection)
        if (stepsToRetract > 0):
          kill move_thread_han_1633
          stopl(0.5)
          $ 1634 "Until (tool_contact_detection)"
          break
        end
        sleep(1.0E-10)
        if (move_thread_flag_1633 > 1):
          join move_thread_han_1633
          break
        end
        sync()
      end
      $ 1635 "Force"
      sleep(0.02)
      zero_ftsensor()
      force_mode(FRM_Reference, [0, 1, 1, 0, 0, 1], [0.0, 0.0, 0.0, 0.0, 0.0, 0.0], 2, [0.1, 0.05, 0.02, 0.3490658503988659, 0.3490658503988659, 3.141592653589793])
      $ 1636 "PSE_T" "noBreak"
      movel(pose_trans(FRM_Reference, PSE_T), a=0.04, v=0.07)
      end_force_mode()
      stopl(5.0)
      $ 1637 "EOAT"
      $ 1638 "rq_move_and_wait_mm(GRP_Open_Pos)"
       rq_move_and_wait_mm (GRP_Open_Pos)
      $ 1639 "OBJ_Picked≔rq_is_object_detected()"
      global OBJ_Picked= rq_is_object_detected ()
      $ 1640 "If PSE_R_H≠PSE_Z"
      if (PSE_R_H != PSE_Z):
        $ 1641 "PSE_R" "breakAfter"
        movel(pose_trans(FRM_Reference, PSE_R), a=0.5, v=0.4, r=0.01)
        $ 1642 "PSE_R_H" "breakAfter"
        movel(pose_trans(FRM_Reference, PSE_R_H), a=0.5, v=0.4)
      else:
        $ 1643 "Else" "noBreak"
        $ 1644 "PSE_R" "breakAfter"
        movel(pose_trans(FRM_Reference, PSE_R), a=0.5, v=0.4)
      end
    elif (8 == switch_1):
      $ 1645 "Case 8"
      $ 1646 "Unload"
      $ 1647 "Action_Info≔'pick object'"
      global Action_Info="pick object"
      $ 1648 "do_transition(pose_trans(FRM_Reference, PSE_T), keep_rxry=OBJ_Picked)"
      do_transition( pose_trans (FRM_Reference, PSE_T), keep_rxry=OBJ_Picked)
      $ 1649 "EOAT"
      $ 1650 "If  not OBJ_Picked"
      if (  not  OBJ_Picked):
        $ 1651 "rq_move_and_wait_mm(GRP_Open_Pos)"
         rq_move_and_wait_mm (GRP_Open_Pos)
      end
      $ 1652 "If PSE_A_H≠PSE_Z"
      if (PSE_A_H != PSE_Z):
        $ 1653 "If JNT_Q≠JNT_Z"
        if (JNT_Q != JNT_Z):
          $ 1654 "movej(get_inverse_kin(pose_trans(FRM_Reference, PSE_A_H), qnear=JNT_Q), r=0.050)"
          movej(get_inverse_kin( pose_trans (FRM_Reference, PSE_A_H), qnear=JNT_Q), r=0.050)
        else:
          $ 1655 "Else" "noBreak"
          $ 1656 "movej(pose_trans(FRM_Reference, PSE_A_H), r=0.050)"
          movej( pose_trans (FRM_Reference, PSE_A_H), r=0.050)
        end
      end
      $ 1657 "If PSE_A≠PSE_Z"
      if (PSE_A != PSE_Z):
        $ 1658 "If JNT_Q≠JNT_Z"
        if (JNT_Q != JNT_Z):
          $ 1659 "movej(get_inverse_kin(pose_trans(FRM_Reference, PSE_A), qnear=JNT_Q), r=0.020)"
          movej(get_inverse_kin( pose_trans (FRM_Reference, PSE_A), qnear=JNT_Q), r=0.020)
        else:
          $ 1660 "Else" "noBreak"
          $ 1661 "movej(pose_trans(FRM_Reference, PSE_A), r=0.020)"
          movej( pose_trans (FRM_Reference, PSE_A), r=0.020)
        end
      end
      $ 1662 "MoveL"
      $ 1663 "If PSE_T_H≠PSE_Z"
      if (PSE_T_H != PSE_Z):
        $ 1664 "PSE_T_H" "breakAfter"
        movel(pose_trans(FRM_Reference, PSE_T_H), a=0.5, v=0.4, r=0.01)
      end
      $ 1665 "PSE_T" "breakAfter"
      movel(pose_trans(FRM_Reference, PSE_T), a=0.08, v=0.12)
      $ 1666 "Force"
      sleep(0.02)
      zero_ftsensor()
      force_mode(FRM_Reference, [1, 1, 0, 0, 0, 0], [0.0, 0.0, 0.0, 0.0, 0.0, 0.0], 2, [0.05, 0.05, 0.1, 0.3490658503988659, 0.3490658503988659, 0.3490658503988659])
      $ 1667 "EOAT" "noBreak"
      $ 1668 "rq_set_force_norm(50)" "noBreak"
       rq_set_force_norm (50)
      $ 1669 "rq_close_and_wait()" "noBreak"
       rq_close_and_wait ()
      $ 1670 "OBJ_Picked≔rq_is_object_detected()" "noBreak"
      global OBJ_Picked= rq_is_object_detected ()
      $ 1671 "If  not OBJ_Picked" "noBreak"
      if (  not  OBJ_Picked):
        $ 1672 "set_error(ERROR_NO_OBJECT_TO_PICK)" "noBreak"
        set_error(ERROR_NO_OBJECT_TO_PICK)
      end
      $ 1673 "If PSE_R_H≠PSE_Z" "noBreak"
      if (PSE_R_H != PSE_Z):
        $ 1674 "PSE_R" "noBreak"
        movel(pose_trans(FRM_Reference, PSE_R), a=0.5, v=0.4, r=0.01)
        $ 1675 "PSE_R_H" "noBreak"
        movel(pose_trans(FRM_Reference, PSE_R_H), a=0.5, v=0.4)
      else:
        $ 1676 "Else" "noBreak"
        $ 1677 "PSE_R" "noBreak"
        movel(pose_trans(FRM_Reference, PSE_R), a=0.5, v=0.4)
      end
      end_force_mode()
      stopl(5.0)
    elif (11 == switch_1):
      $ 1678 "Case 11"
      $ 1679 "Place without opening gripper"
      $ 1680 "Action_Info≔'place object without gripper opening'"
      global Action_Info="place object without gripper opening"
      $ 1682 "movel(FRM_Container_S, a=0.025, v=0.015, r=0.00001)"
      movel(FRM_Container_S, a=0.025, v=0.015, r=0.00001)
      $ 1683 "EXTT"
      $ 1684 "Switch JIG"
      switch_2 = JIG
      $ 1685 "Case 1"
      if (1 == switch_2):
        $ 1686 "3FG"
        $ 1687 "If OBJ_Picked"
        if (OBJ_Picked):
          $ 1688 "Set GRP_3F_Open=On"
          set_standard_digital_out(5, True)
        end
      end
      $ 1689 "If PSE_A_H≠PSE_Z"
      if (PSE_A_H != PSE_Z):
        $ 1690 "If JNT_Q≠JNT_Z"
        if (JNT_Q != JNT_Z):
          $ 1691 "movej(get_inverse_kin(pose_trans(FRM_Reference, PSE_A_H), qnear=JNT_Q), r=0.050)"
          movej(get_inverse_kin( pose_trans (FRM_Reference, PSE_A_H), qnear=JNT_Q), r=0.050)
        else:
          $ 1692 "Else" "noBreak"
          $ 1693 "movej(pose_trans(FRM_Reference, PSE_A_H), r=0.050)"
          movej( pose_trans (FRM_Reference, PSE_A_H), r=0.050)
        end
      end
      $ 1694 "If PSE_A≠PSE_Z"
      if (PSE_A != PSE_Z):
        $ 1695 "If JNT_Q≠JNT_Z"
        if (JNT_Q != JNT_Z):
          $ 1696 "movej(get_inverse_kin(pose_trans(FRM_Reference, PSE_A), qnear=JNT_Q), r=0.020)"
          movej(get_inverse_kin( pose_trans (FRM_Reference, PSE_A), qnear=JNT_Q), r=0.020)
        else:
          $ 1697 "Else" "noBreak"
          $ 1698 "movej(pose_trans(FRM_Reference, PSE_A), r=0.020)"
          movej( pose_trans (FRM_Reference, PSE_A), r=0.020)
        end
      end
      $ 1699 "MoveL"
      $ 1700 "If PSE_T_H≠PSE_Z"
      if (PSE_T_H != PSE_Z):
        $ 1701 "PSE_T_H" "breakAfter"
        movel(pose_trans(FRM_Reference, PSE_T_H), a=0.5, v=0.4, r=0.01)
      end
      $ 1702 "PSE_T" "breakAfter"
      global move_thread_flag_1702=0
      thread move_thread_1702():
        enter_critical
        move_thread_flag_1702 = 1
        movel(pose_trans(FRM_Reference, PSE_T), a=0.05, v=0.09)
        move_thread_flag_1702 = 2
        exit_critical
      end
      move_thread_flag_1702 = 0
      move_thread_han_1702 = run move_thread_1702()
      while (True):
        local targetTcpDirection=get_target_tcp_speed()
        local stepsToRetract=tool_contact(direction=targetTcpDirection)
        if (stepsToRetract > 0):
          kill move_thread_han_1702
          stopl(0.5)
          $ 1703 "Until (tool_contact_detection)"
          break
        end
        sleep(1.0E-10)
        if (move_thread_flag_1702 > 1):
          join move_thread_han_1702
          break
        end
        sync()
      end
      $ 1704 "Force"
      sleep(0.02)
      zero_ftsensor()
      force_mode(FRM_Reference, [1, 1, 1, 0, 0, 0], [0.0, 0.0, 0.0, 0.0, 0.0, 0.0], 2, [0.1, 0.1, 0.01, 0.3490658503988659, 0.3490658503988659, 0.3490658503988659])
      $ 1705 "PSE_T" "noBreak"
      movel(pose_trans(FRM_Reference, PSE_T), a=0.04, v=0.07)
      end_force_mode()
      stopl(5.0)
      $ 1706 "EXTT"
      $ 1707 "Switch JIG"
      switch_2 = JIG
      $ 1708 "Case 1"
      if (1 == switch_2):
        $ 1709 "3FG"
        $ 1710 "If OBJ_Picked"
        if (OBJ_Picked):
          $ 1711 "Set GRP_3F_Open=Off"
          set_standard_digital_out(5, False)
          $ 1712 "Wait: 0.2"
          sleep(0.2)
        end
      end
      $ 1713 "EOAT"
      $ 1714 "Comment"
      # Comment
    elif (12 == switch_1):
      $ 1715 "Case 12"
      $ 1716 "Decap"
      $ 1717 "Action_Info≔'decapping'"
      global Action_Info="decapping"
      $ 1718 "Set GRP_3F_Enable=On"
      set_standard_digital_out(4, True)
      $ 1719 "Set GRP_3F_Decap=On"
      set_standard_digital_out(3, True)
      $ 1720 "Force"
      sleep(0.02)
      zero_ftsensor()
      force_mode(tool_pose(), [0, 0, 1, 0, 0, 0], [0.0, 0.0, 5.0, 0.0, 0.0, 0.0], 2, [0.1, 0.1, 0.15, 0.3490658503988659, 0.3490658503988659, 0.3490658503988659])
      $ 1721 "check_decapping(offset=0.015, timeout=5, abort=CMD_Hold)" "noBreak"
      check_decapping(offset=0.015, timeout=5, abort=CMD_Hold)
      end_force_mode()
      stopl(5.0)
      $ 1722 "Set GRP_3F_Decap=Off"
      set_standard_digital_out(3, False)
      $ 1723 "Set GRP_3F_Enable=Off"
      set_standard_digital_out(4, False)
      $ 1724 "MoveL"
      $ 1725 "PSE_R" "breakAfter"
      movel(pose_trans(FRM_Reference, PSE_R), a=0.8, v=0.15)
    elif (13 == switch_1):
      $ 1726 "Case 13"
      $ 1727 "TMR_Barcode: Reset"
      TMR_Barcode = 0
      $ 1728 "Read"
      $ 1729 "TMR_Barcode: Start"
      TMR_Barcode_is_counting = True
      $ 1730 "If TMR_Barcode<PRM_TO_Read_BC"
      global thread_flag_1730=0
      thread Thread_if_1730():
        $ 1731 "KeyenceTrigger"
        $ 1732 "Set OClearResult=HI:Pulse 0.2"
        thread SinglePulse2():
          write_output_boolean_register(2, True)
          sleep(0.2)
          write_output_boolean_register(2, False)
        end
        singlePulse2 = run SinglePulse2()
        $ 1733 "Wait: 0.5"
        sleep(0.5)
        $ 1734 "Set OTriggerBarcode=Off"
        write_output_boolean_register(1, False)
        $ 1735 "Wait: 0.5"
        sleep(0.5)
        $ 1736 "Set OTriggerBarcode=On"
        write_output_boolean_register(1, True)
        $ 1737 "Wait: 0.5"
        sleep(0.5)
        $ 1738 "Preorient"
        $ 1739 "TMR_Barcode: Reset"
        TMR_Barcode = 0
        $ 1740 "If ICmdExctd"
        if (read_input_boolean_register(12)):
          $ 1741 "Set GRP_3F_Decap=On"
          set_standard_digital_out(3, True)
          $ 1742 "Set GRP_3F_Enable=On"
          set_standard_digital_out(4, True)
          $ 1743 "Loop ICmdExctd"
          while (read_input_boolean_register(12)):
            $ 1744 "KeyenceTrigger"
            $ 1745 "Set OClearResult=HI:Pulse 0.1"
            thread SinglePulse3():
              write_output_boolean_register(2, True)
              sleep(0.1)
              write_output_boolean_register(2, False)
            end
            singlePulse3 = run SinglePulse3()
            $ 1746 "Wait: 0.3"
            sleep(0.3)
            $ 1747 "Set OTriggerBarcode=Off"
            write_output_boolean_register(1, False)
            $ 1748 "Wait: 0.3"
            sleep(0.3)
            $ 1749 "Set OTriggerBarcode=On"
            write_output_boolean_register(1, True)
            $ 1750 "Wait: 0.1"
            sleep(0.1)
          end
        end
        $ 1751 "If  not ICmdExctd"
        if (  not  read_input_boolean_register(12)):
          $ 1752 "Set GRP_3F_Decap=On"
          set_standard_digital_out(3, True)
          $ 1753 "Set GRP_3F_Enable=On"
          set_standard_digital_out(4, True)
          $ 1754 "Wait ICmdExctd=HI"
          while (read_input_boolean_register(12) == False):
            sync()
          end
        end
        $ 1755 "Set GRP_3F_Decap=Off"
        set_standard_digital_out(3, False)
        $ 1756 "Set GRP_3F_Enable=Off"
        set_standard_digital_out(4, False)
        $ 1757 "OBJ_Brc_OK≔ True "
        global OBJ_Brc_OK=  True
        thread_flag_1730 = 1
      end
      if (TMR_Barcode<PRM_TO_Read_BC):
        global thread_handler_1730=run Thread_if_1730()
        while (thread_flag_1730 == 0):
          if not(TMR_Barcode<PRM_TO_Read_BC):
            kill thread_handler_1730
            thread_flag_1730 = 2
          else:
            sync()
          end
        end
      else:
        thread_flag_1730 = 2
      end
      if (thread_flag_1730 == 2):
        $ 1758 "Else" "noBreak"
        $ 1759 "exeption"
        $ 1760 "error"
        $ 1762 "OBJ_Brc_OK≔ False "
        global OBJ_Brc_OK=  False
      end
      $ 1763 "Set GRP_3F_Decap=Off"
      set_standard_digital_out(3, False)
      $ 1764 "Set GRP_3F_Enable=Off"
      set_standard_digital_out(4, False)
      $ 1765 "Set OTriggerBarcode=Off"
      write_output_boolean_register(1, False)
    elif (15 == switch_1):
      $ 1766 "Case 15"
      $ 1767 "Detect"
      $ 1768 "Action_Info≔'detect'"
      global Action_Info="detect"
    elif (30 == switch_1):
      $ 1769 "Case 30"
      $ 1770 "Shake"
      $ 1771 "Action_Info≔'shake'"
      global Action_Info="shake"
      $ 1772 "do_transition(pose_trans(FRM_Reference, PSE_T), keep_rxry=OBJ_Picked)"
      do_transition( pose_trans (FRM_Reference, PSE_T), keep_rxry=OBJ_Picked)
      $ 1773 "If PSE_A_H≠PSE_Z"
      if (PSE_A_H != PSE_Z):
        $ 1774 "If JNT_Q≠JNT_Z"
        if (JNT_Q != JNT_Z):
          $ 1775 "movej(get_inverse_kin(pose_trans(FRM_Reference, PSE_A_H), qnear=JNT_Q), r=0.050)"
          movej(get_inverse_kin( pose_trans (FRM_Reference, PSE_A_H), qnear=JNT_Q), r=0.050)
        else:
          $ 1776 "Else" "noBreak"
          $ 1777 "movej(pose_trans(FRM_Reference, PSE_A_H), r=0.050)"
          movej( pose_trans (FRM_Reference, PSE_A_H), r=0.050)
        end
      end
      $ 1778 "If PSE_A≠PSE_Z"
      if (PSE_A != PSE_Z):
        $ 1779 "If JNT_Q≠JNT_Z"
        if (JNT_Q != JNT_Z):
          $ 1780 "movej(get_inverse_kin(pose_trans(FRM_Reference, PSE_A), qnear=JNT_Q), r=0.020)"
          movej(get_inverse_kin( pose_trans (FRM_Reference, PSE_A), qnear=JNT_Q), r=0.020)
        else:
          $ 1781 "Else" "noBreak"
          $ 1782 "movej(pose_trans(FRM_Reference, PSE_A), r=0.020)"
          movej( pose_trans (FRM_Reference, PSE_A), r=0.020)
        end
      end
      $ 1783 "MoveL"
      $ 1784 "If PSE_T_H≠PSE_Z"
      if (PSE_T_H != PSE_Z):
        $ 1785 "PSE_T_H" "breakAfter"
        movel(pose_trans(FRM_Reference, PSE_T_H), a=0.5, v=0.4, r=0.01)
      end
      $ 1786 "PSE_T" "breakAfter"
      movel(pose_trans(FRM_Reference, PSE_T), a=0.08, v=0.12)
      $ 1787 "EXTT"
      $ 1788 "Comment"
      # Comment
      $ 1789 "MoveJ"
      $ 1790 "Waypoint_6" "breakAfter"
      movej(get_inverse_kin(Waypoint_6_p, qnear=Waypoint_6_q), a=1.3962634015954636, v=1.0471975511965976)
      $ 1791 "MoveJ"
      $ 1792 "Waypoint_18" "breakAfter"
      movej(get_inverse_kin(Waypoint_18_p, qnear=Waypoint_18_q), a=1.3962634015954636, v=1.0471975511965976)
      $ 1793 "MoveJ"
      $ 1794 "Waypoint_12" "breakAfter"
      movej(get_inverse_kin(Waypoint_12_p, qnear=Waypoint_12_q), a=1.3962634015954636, v=1.0471975511965976)
      $ 1795 "MoveJ"
      $ 1796 "Waypoint_19" "breakAfter"
      movej(get_inverse_kin(Waypoint_19_p, qnear=Waypoint_19_q), a=1.3962634015954636, v=1.0471975511965976)
      $ 1797 "If PSE_R_H≠PSE_Z"
      if (PSE_R_H != PSE_Z):
        $ 1798 "PSE_R" "breakAfter"
        movel(pose_trans(FRM_Reference, PSE_R), a=0.5, v=0.4, r=0.01)
        $ 1799 "PSE_R_H" "breakAfter"
        movel(pose_trans(FRM_Reference, PSE_R_H), a=0.5, v=0.4)
      else:
        $ 1800 "Else" "noBreak"
        $ 1801 "PSE_R" "breakAfter"
        movel(pose_trans(FRM_Reference, PSE_R), a=0.5, v=0.4)
      end
    elif (31 == switch_1):
      $ 1802 "Case 31"
      $ 1803 "Action_Info≔'Pick_Vial'"
      global Action_Info="Pick_Vial"
      $ 1804 "Pick_Vial"
      # begin: URCap Program Node
      #   Source: Robotiq_Grippers, 1.8.4.4844, Robotiq Inc.
      #   Type: Gripper
      $ 1805 "Gripper Open (1)"
      if not(gripper_connected[0]):
        popup("Gripper 1 must be connected to run this program.", "No connection", False, True, True)
      end
      if not(rq_is_gripper_activated("1")):
        popup("Gripper 1 is not activated. Go to Installation tab > Gripper to activate it and run the program again.", "Not activated", False, True, True)
      end
      rq_set_pos_spd_for(0, 82, 71, "1")
      rq_wait_pos_spe_for_request(0, 82, 71, "1")
      rq_go_to("1")
      rq_wait("1")
      # end: URCap Program Node
      $ 1806 "MoveJ"
      $ 1807 "Vial_above" "breakAfter"
      movej(get_inverse_kin(Vial_above_p, qnear=Vial_above_q), a=0.5235987755982988, v=0.4363323129985824, r=0.05)
      $ 1808 "MoveL"
      $ 1809 "Vial_pick_point" "breakAfter"
      movel(Vial_pick_point_p, a=0.5, v=0.1)
      # begin: URCap Program Node
      #   Source: Robotiq_Grippers, 1.8.4.4844, Robotiq Inc.
      #   Type: Gripper
      $ 1810 "Gripper Close (1)"
      if not(gripper_connected[0]):
        popup("Gripper 1 must be connected to run this program.", "No connection", False, True, True)
      end
      if not(rq_is_gripper_activated("1")):
        popup("Gripper 1 is not activated. Go to Installation tab > Gripper to activate it and run the program again.", "Not activated", False, True, True)
      end
      rq_set_pos_spd_for(255, 71, 84, "1")
      rq_wait_pos_spe_for_request(255, 71, 84, "1")
      rq_go_to("1")
      rq_wait("1")
      # end: URCap Program Node
      $ 1811 "MoveL"
      $ 1812 "Waypoint_20" "breakAfter"
      movel(Waypoint_20_p, a=0.5, v=0.1, r=0.05)
      $ 1813 "Home (Safe)"
      movej([-1.2302089344500047, -1.2969853503591224, -1.875639182904262, -1.539621866126728, 1.5731943360401213, -2.80099559440227], a=1.3962634015954636, v=1.0471975511965976)
    elif (32 == switch_1):
      $ 1814 "Case 32"
      $ 1815 "decap≔ False "
      global decap=  False
      $ 1816 "decap_Vial"
      $ 1817 "Set GRP_3F_Open=On"
      set_standard_digital_out(5, True)
      $ 1818 "MoveJ"
      $ 1819 "Waypoint_33" "breakAfter"
      movej(get_inverse_kin(Waypoint_33_p, qnear=Waypoint_33_q), a=0.5235987755982988, v=0.4363323129985824)
      $ 1820 "MoveL"
      $ 1821 "Vial_3FG_place" "breakAfter"
      movel(Vial_3FG_place_p, a=0.5, v=0.1)
      $ 1822 "Set GRP_3F_Open=Off"
      set_standard_digital_out(5, False)
      $ 1823 "Wait: 0.5"
      sleep(0.5)
      $ 1824 "MoveL"
      $ 1825 "Waypoint_34" "breakAfter"
      movel(Waypoint_34_p, a=0.5, v=0.1, r=0.05)
      $ 1826 "MoveJ"
      $ 1827 "cap_dump" "breakAfter"
      movej(get_inverse_kin(cap_dump_p, qnear=cap_dump_q), a=0.5235987755982988, v=0.4363323129985824)
      # begin: URCap Program Node
      #   Source: Robotiq_Grippers, 1.8.4.4844, Robotiq Inc.
      #   Type: Gripper
      $ 1828 "Gripper Open (1)"
      if not(gripper_connected[0]):
        popup("Gripper 1 must be connected to run this program.", "No connection", False, True, True)
      end
      if not(rq_is_gripper_activated("1")):
        popup("Gripper 1 is not activated. Go to Installation tab > Gripper to activate it and run the program again.", "Not activated", False, True, True)
      end
      rq_set_pos_spd_for(0, 255, 255, "1")
      rq_wait_pos_spe_for_request(0, 255, 255, "1")
      rq_go_to("1")
      rq_wait("1")
      # end: URCap Program Node
      $ 1829 "MoveJ"
      $ 1830 "Waypoint_35" "breakAfter"
      movej(get_inverse_kin(Waypoint_35_p, qnear=Waypoint_35_q), a=0.5235987755982988, v=0.4363323129985824, r=0.05)
      $ 1831 "MoveL"
      $ 1832 "Vial_3FG_place" "breakAfter"
      movel(Vial_3FG_place_p, a=0.5, v=0.1)
      # begin: URCap Program Node
      #   Source: Robotiq_Grippers, 1.8.4.4844, Robotiq Inc.
      #   Type: Gripper
      $ 1833 "Gripper Close (1)"
      if not(gripper_connected[0]):
        popup("Gripper 1 must be connected to run this program.", "No connection", False, True, True)
      end
      if not(rq_is_gripper_activated("1")):
        popup("Gripper 1 is not activated. Go to Installation tab > Gripper to activate it and run the program again.", "Not activated", False, True, True)
      end
      rq_set_pos_spd_for(255, 204, 255, "1")
      rq_wait_pos_spe_for_request(255, 204, 255, "1")
      rq_go_to("1")
      rq_wait("1")
      # end: URCap Program Node
      $ 1840 "Decap"
      $ 1841 "Action_Info≔'decapping'"
      global Action_Info="decapping"
      $ 1842 "Set GRP_3F_Enable=On"
      set_standard_digital_out(4, True)
      $ 1843 "Set GRP_3F_Decap=On"
      set_standard_digital_out(3, True)
      $ 1844 "Force"
      sleep(0.02)
      zero_ftsensor()
      force_mode(p[0.0,0.0,0.0,0.0,0.0,0.0], [0, 0, 1, 0, 0, 0], [0.0, 0.0, 1.0, 0.0, 0.0, 0.0], 2, [0.1, 0.1, 0.001, 0.3490658503988659, 0.3490658503988659, 0.3490658503988659])
      $ 1845 "check_decapping(offset=0.015, timeout=10, abort=CMD_Hold)" "noBreak"
      check_decapping(offset=0.015, timeout=10, abort=CMD_Hold)
      end_force_mode()
      stopl(5.0)
      $ 1846 "Set GRP_3F_Decap=Off"
      set_standard_digital_out(3, False)
      $ 1847 "Set GRP_3F_Enable=Off"
      set_standard_digital_out(4, False)
      $ 1848 "MoveL"
      $ 1849 "Waypoint_36" "breakAfter"
      movel(Waypoint_36_p, a=0.5, v=0.1, r=0.05)
      $ 1850 "MoveJ"
      $ 1851 "cap_dump" "breakAfter"
      movej(get_inverse_kin(cap_dump_p, qnear=cap_dump_q), a=0.5235987755982988, v=0.4363323129985824)
      # begin: URCap Program Node
      #   Source: Robotiq_Grippers, 1.8.4.4844, Robotiq Inc.
      #   Type: Gripper
      $ 1852 "Gripper Open (1)"
      if not(gripper_connected[0]):
        popup("Gripper 1 must be connected to run this program.", "No connection", False, True, True)
      end
      if not(rq_is_gripper_activated("1")):
